Universal Robots URScript: FaiChun_9 Jan_4.script

def Machining1():
  # Default parameters:
  global speed_ms = 0.3
  global speed_rads = 0.75
  global accel_mss = 3
  global accel_radss = 1.2
  global blend_radius_m = 0.0003

  # Add subprograms here
  # Start of main program
  # Program generated by RoboDK v5.6.8 for UR10e on 09/01/2025 17:05:57
  # Using nominal kinematics.
  blend_radius_m = 0.0003
  speed_ms = 0.03
  # set_reference(p[0.335000, -0.060000, 0.000000, 0.000000, 0.000000, 0.000000])
  set_tcp(p[0.000000, 0.000000, 0.252000, 0.000000, 0.000000, 0.000000])
  # Show Tool
  movej([0.372931, -1.100475, -2.621390, -0.990524, 1.570796, 1.943727],accel_radss,speed_rads,0,blend_radius_m)
  movel([0.372931, -1.160560, -2.660288, -0.891541, 1.570796, 1.943727],accel_mss,speed_ms,0,blend_radius_m)
  #SetTool1
  #M_RunCode6
  #SetRPM60000
  speed_ms = 0.03
  #M_RunCode3
  movel([0.372931, -1.188229, -2.675077, -0.849084, 1.570796, 1.943727],accel_mss,speed_ms,0,blend_radius_m)
  speed_ms = 0.003
  movel([0.372931, -1.195517, -2.678710, -0.838162, 1.570796, 1.943727],accel_mss,speed_ms,0,blend_radius_m)
  speed_ms = 0.007
  movel([0.375174, -1.198382, -2.677355, -0.836652, 1.570796, 1.945970],accel_mss,speed_ms,0,blend_radius_m)
  movel([0.377606, -1.200493, -2.676351, -0.835545, 1.570796, 1.948402],accel_mss,speed_ms,0,blend_radius_m)
  movel([0.380241, -1.201847, -2.675704, -0.834837, 1.570796, 1.951037],accel_mss,speed_ms,0,blend_radius_m)
  movel([0.383075, -1.202452, -2.675415, -0.834522, 1.570796, 1.953872],accel_mss,speed_ms,0,blend_radius_m)
  movel([0.386053, -1.202396, -2.675442, -0.834551, 1.570796, 1.956849],accel_mss,speed_ms,0,blend_radius_m)
  movel([0.389105, -1.201761, -2.675746, -0.834882, 1.570796, 1.959901],accel_mss,speed_ms,0,blend_radius_m)
  movel([0.392242, -1.200547, -2.676325, -0.835516, 1.570796, 1.963038],accel_mss,speed_ms,0,blend_radius_m)
  movel([0.395468, -1.198746, -2.677183, -0.836461, 1.570796, 1.966265],accel_mss,speed_ms,0,blend_radius_m)
  movel([0.380728, -1.210997, -2.671282, -0.830110, 1.570796, 1.951524],accel_mss,speed_ms,0,blend_radius_m)
  movel([0.361187, -1.181602, -2.685164, -0.845623, 1.570796, 1.931983],accel_mss,speed_ms,0,blend_radius_m)
  movel([0.362683, -1.180288, -2.685763, -0.846338, 1.570796, 1.933479],accel_mss,speed_ms,0,blend_radius_m)
  movel([0.366731, -1.177285, -2.687125, -0.847980, 1.570796, 1.937528],accel_mss,speed_ms,0,blend_radius_m)
  movel([0.371187, -1.175024, -2.688143, -0.849221, 1.570796, 1.941984],accel_mss,speed_ms,0,blend_radius_m)
  movel([0.375796, -1.173412, -2.688867, -0.850111, 1.570796, 1.946593],accel_mss,speed_ms,0,blend_radius_m)
  movel([0.380308, -1.172343, -2.689344, -0.850701, 1.570796, 1.951104],accel_mss,speed_ms,0,blend_radius_m)
  movel([0.392053, -1.170737, -2.690060, -0.851592, 1.570796, 1.962849],accel_mss,speed_ms,0,blend_radius_m)
  movel([0.402871, -1.169477, -2.690620, -0.852292, 1.570796, 1.973667],accel_mss,speed_ms,0,blend_radius_m)
  movel([0.407062, -1.168614, -2.691003, -0.852772, 1.570796, 1.977858],accel_mss,speed_ms,0,blend_radius_m)
  movel([0.411263, -1.167290, -2.691588, -0.853511, 1.570796, 1.982060],accel_mss,speed_ms,0,blend_radius_m)
  movel([0.415272, -1.165416, -2.692413, -0.854560, 1.570796, 1.986068],accel_mss,speed_ms,0,blend_radius_m)
  movel([0.418891, -1.162891, -2.693519, -0.855978, 1.570796, 1.989688],accel_mss,speed_ms,0,blend_radius_m)
  movel([0.422708, -1.159075, -2.695179, -0.858136, 1.570796, 1.993505],accel_mss,speed_ms,0,blend_radius_m)
  movel([0.424029, -1.157173, -2.696000, -0.859216, 1.570796, 1.994826],accel_mss,speed_ms,0,blend_radius_m)
  movel([0.424957, -1.155274, -2.696817, -0.860298, 1.570796, 1.995753],accel_mss,speed_ms,0,blend_radius_m)
  movel([0.425724, -1.151821, -2.698292, -0.862276, 1.570796, 1.996520],accel_mss,speed_ms,0,blend_radius_m)
  movel([0.425106, -1.149060, -2.699463, -0.863866, 1.570796, 1.995903],accel_mss,speed_ms,0,blend_radius_m)
  movel([0.424036, -1.147738, -2.700021, -0.864630, 1.570796, 1.994833],accel_mss,speed_ms,0,blend_radius_m)
  movel([0.422706, -1.147211, -2.700243, -0.864935, 1.570796, 1.993503],accel_mss,speed_ms,0,blend_radius_m)
  movel([0.421264, -1.147406, -2.700161, -0.864822, 1.570796, 1.992060],accel_mss,speed_ms,0,blend_radius_m)
  movel([0.419851, -1.148255, -2.699803, -0.864331, 1.570796, 1.990647],accel_mss,speed_ms,0,blend_radius_m)
  movel([0.418269, -1.150392, -2.698899, -0.863098, 1.570796, 1.989065],accel_mss,speed_ms,0,blend_radius_m)
  movel([0.416848, -1.152543, -2.697985, -0.861862, 1.570796, 1.987644],accel_mss,speed_ms,0,blend_radius_m)
  movel([0.414611, -1.154776, -2.697030, -0.860583, 1.570796, 1.985407],accel_mss,speed_ms,0,blend_radius_m)
  movel([0.411600, -1.156758, -2.696179, -0.859452, 1.570796, 1.982396],accel_mss,speed_ms,0,blend_radius_m)
  movel([0.408872, -1.157382, -2.695910, -0.859097, 1.570796, 1.979668],accel_mss,speed_ms,0,blend_radius_m)
  movel([0.406625, -1.156830, -2.696148, -0.859411, 1.570796, 1.977422],accel_mss,speed_ms,0,blend_radius_m)
  movel([0.405066, -1.155270, -2.696818, -0.860301, 1.570796, 1.975862],accel_mss,speed_ms,0,blend_radius_m)
  movel([0.404360, -1.152976, -2.697800, -0.861613, 1.570796, 1.975156],accel_mss,speed_ms,0,blend_radius_m)
  movel([0.404684, -1.150222, -2.698971, -0.863196, 1.570796, 1.975481],accel_mss,speed_ms,0,blend_radius_m)
  movel([0.406108, -1.147296, -2.700207, -0.864886, 1.570796, 1.976904],accel_mss,speed_ms,0,blend_radius_m)
  movel([0.408704, -1.144500, -2.701381, -0.866509, 1.570796, 1.979501],accel_mss,speed_ms,0,blend_radius_m)
  movel([0.411321, -1.142589, -2.702178, -0.867622, 1.570796, 1.982118],accel_mss,speed_ms,0,blend_radius_m)
  movel([0.413891, -1.141382, -2.702680, -0.868328, 1.570796, 1.984688],accel_mss,speed_ms,0,blend_radius_m)
  movel([0.416415, -1.140882, -2.702887, -0.868620, 1.570796, 1.987211],accel_mss,speed_ms,0,blend_radius_m)
  movel([0.418874, -1.141102, -2.702796, -0.868491, 1.570796, 1.989670],accel_mss,speed_ms,0,blend_radius_m)
  movel([0.421187, -1.141949, -2.702444, -0.867996, 1.570796, 1.991984],accel_mss,speed_ms,0,blend_radius_m)
  movel([0.423263, -1.143337, -2.701866, -0.867186, 1.570796, 1.994060],accel_mss,speed_ms,0,blend_radius_m)
  movel([0.426702, -1.147727, -2.700026, -0.864636, 1.570796, 1.997499],accel_mss,speed_ms,0,blend_radius_m)
  movel([0.428202, -1.151149, -2.698578, -0.862662, 1.570796, 1.998999],accel_mss,speed_ms,0,blend_radius_m)
  movel([0.429111, -1.154788, -2.697025, -0.860576, 1.570796, 1.999907],accel_mss,speed_ms,0,blend_radius_m)
  movel([0.429435, -1.158639, -2.695367, -0.858383, 1.570796, 2.000231],accel_mss,speed_ms,0,blend_radius_m)
  movel([0.429184, -1.162688, -2.693608, -0.856093, 1.570796, 1.999980],accel_mss,speed_ms,0,blend_radius_m)
  movel([0.428147, -1.166773, -2.691816, -0.853800, 1.570796, 1.998944],accel_mss,speed_ms,0,blend_radius_m)
  movel([0.426123, -1.170732, -2.690063, -0.851595, 1.570796, 1.996919],accel_mss,speed_ms,0,blend_radius_m)
  movel([0.423112, -1.174570, -2.688347, -0.849472, 1.570796, 1.993908],accel_mss,speed_ms,0,blend_radius_m)
  movel([0.419124, -1.178294, -2.686668, -0.847427, 1.570796, 1.989921],accel_mss,speed_ms,0,blend_radius_m)
  movel([0.415165, -1.181134, -2.685378, -0.845877, 1.570796, 1.985962],accel_mss,speed_ms,0,blend_radius_m)
  movel([0.411168, -1.183199, -2.684434, -0.844756, 1.570796, 1.981965],accel_mss,speed_ms,0,blend_radius_m)
  movel([0.407228, -1.184627, -2.683779, -0.843983, 1.570796, 1.978024],accel_mss,speed_ms,0,blend_radius_m)
  movel([0.403450, -1.185553, -2.683353, -0.843483, 1.570796, 1.974246],accel_mss,speed_ms,0,blend_radius_m)
  movel([0.394479, -1.186696, -2.682826, -0.842867, 1.570796, 1.965275],accel_mss,speed_ms,0,blend_radius_m)
  movel([0.385975, -1.187888, -2.682274, -0.842226, 1.570796, 1.956771],accel_mss,speed_ms,0,blend_radius_m)
  movel([0.382534, -1.188768, -2.681867, -0.841754, 1.570796, 1.953330],accel_mss,speed_ms,0,blend_radius_m)
  movel([0.379011, -1.190092, -2.681251, -0.841046, 1.570796, 1.949807],accel_mss,speed_ms,0,blend_radius_m)
  movel([0.375525, -1.191944, -2.680387, -0.840058, 1.570796, 1.946321],accel_mss,speed_ms,0,blend_radius_m)
  movel([0.372203, -1.194411, -2.679231, -0.838747, 1.570796, 1.942999],accel_mss,speed_ms,0,blend_radius_m)
  movel([0.372931, -1.195517, -2.678710, -0.838162, 1.570796, 1.943727],accel_mss,speed_ms,0,blend_radius_m)
  speed_ms = 0.003
  movel([0.372931, -1.188229, -2.675077, -0.849084, 1.570796, 1.943727],accel_mss,speed_ms,0,blend_radius_m)
  speed_ms = 0.03
  movel([0.372931, -1.160560, -2.660288, -0.891541, 1.570796, 1.943727],accel_mss,speed_ms,0,blend_radius_m)
  #M_RunCode9
  movel([0.396562, -1.185032, -2.648957, -0.878400, 1.570796, 1.967359],accel_mss,speed_ms,0,blend_radius_m)
  #M_RunCode3
  movel([0.396562, -1.212507, -2.663422, -0.836459, 1.570796, 1.967359],accel_mss,speed_ms,0,blend_radius_m)
  speed_ms = 0.003
  movel([0.396562, -1.219730, -2.666973, -0.825686, 1.570796, 1.967359],accel_mss,speed_ms,0,blend_radius_m)
  speed_ms = 0.007
  movel([0.404177, -1.212524, -2.670535, -0.829330, 1.570796, 1.974973],accel_mss,speed_ms,0,blend_radius_m)
  movel([0.415586, -1.202971, -2.675166, -0.834252, 1.570796, 1.986383],accel_mss,speed_ms,0,blend_radius_m)
  movel([0.427444, -1.193807, -2.679515, -0.839067, 1.570796, 1.998240],accel_mss,speed_ms,0,blend_radius_m)
  movel([0.436211, -1.187874, -2.682281, -0.842234, 1.570796, 2.007007],accel_mss,speed_ms,0,blend_radius_m)
  movel([0.439450, -1.186181, -2.683064, -0.843145, 1.570796, 2.010246],accel_mss,speed_ms,0,blend_radius_m)
  movel([0.441984, -1.185395, -2.683426, -0.843569, 1.570796, 2.012781],accel_mss,speed_ms,0,blend_radius_m)
  movel([0.443806, -1.185518, -2.683369, -0.843502, 1.570796, 2.014603],accel_mss,speed_ms,0,blend_radius_m)
  movel([0.444914, -1.186554, -2.682891, -0.842944, 1.570796, 2.015710],accel_mss,speed_ms,0,blend_radius_m)
  movel([0.445184, -1.188242, -2.682110, -0.842036, 1.570796, 2.015980],accel_mss,speed_ms,0,blend_radius_m)
  movel([0.444497, -1.190341, -2.681135, -0.840912, 1.570796, 2.015293],accel_mss,speed_ms,0,blend_radius_m)
  movel([0.442860, -1.192839, -2.679968, -0.839581, 1.570796, 2.013656],accel_mss,speed_ms,0,blend_radius_m)
  movel([0.440283, -1.195736, -2.678607, -0.838046, 1.570796, 2.011079],accel_mss,speed_ms,0,blend_radius_m)
  movel([0.432369, -1.203009, -2.675148, -0.834232, 1.570796, 2.003165],accel_mss,speed_ms,0,blend_radius_m)
  movel([0.420879, -1.212434, -2.670579, -0.829376, 1.570796, 1.991675],accel_mss,speed_ms,0,blend_radius_m)
  movel([0.409297, -1.221297, -2.666191, -0.824901, 1.570796, 1.980094],accel_mss,speed_ms,0,blend_radius_m)
  movel([0.400914, -1.226977, -2.663332, -0.822080, 1.570796, 1.971711],accel_mss,speed_ms,0,blend_radius_m)
  movel([0.397832, -1.228606, -2.662505, -0.821278, 1.570796, 1.968628],accel_mss,speed_ms,0,blend_radius_m)
  movel([0.395403, -1.229390, -2.662106, -0.820893, 1.570796, 1.966199],accel_mss,speed_ms,0,blend_radius_m)
  movel([0.393621, -1.229327, -2.662138, -0.820924, 1.570796, 1.964417],accel_mss,speed_ms,0,blend_radius_m)
  movel([0.392480, -1.228419, -2.662600, -0.821370, 1.570796, 1.963276],accel_mss,speed_ms,0,blend_radius_m)
  movel([0.392118, -1.226877, -2.663382, -0.822130, 1.570796, 1.962915],accel_mss,speed_ms,0,blend_radius_m)
  movel([0.392674, -1.224917, -2.664373, -0.823099, 1.570796, 1.963470],accel_mss,speed_ms,0,blend_radius_m)
  movel([0.394153, -1.222536, -2.665570, -0.824283, 1.570796, 1.964950],accel_mss,speed_ms,0,blend_radius_m)
  movel([0.396562, -1.219730, -2.666973, -0.825686, 1.570796, 1.967359],accel_mss,speed_ms,0,blend_radius_m)
  speed_ms = 0.003
  movel([0.396562, -1.212507, -2.663422, -0.836459, 1.570796, 1.967359],accel_mss,speed_ms,0,blend_radius_m)
  speed_ms = 0.03
  movel([0.396562, -1.185032, -2.648957, -0.878400, 1.570796, 1.967359],accel_mss,speed_ms,0,blend_radius_m)
  #M_RunCode9
  movel([0.389349, -1.187940, -2.647569, -0.876881, 1.570796, 1.960145],accel_mss,speed_ms,0,blend_radius_m)
  #M_RunCode3
  movel([0.389349, -1.215389, -2.661996, -0.835005, 1.570796, 1.960145],accel_mss,speed_ms,0,blend_radius_m)
  speed_ms = 0.003
  movel([0.389349, -1.222603, -2.665537, -0.824249, 1.570796, 1.960145],accel_mss,speed_ms,0,blend_radius_m)
  speed_ms = 0.007
  movel([0.389682, -1.219825, -2.666926, -0.825638, 1.570796, 1.960478],accel_mss,speed_ms,0,blend_radius_m)
  movel([0.390483, -1.216852, -2.668402, -0.827134, 1.570796, 1.961280],accel_mss,speed_ms,0,blend_radius_m)
  movel([0.391770, -1.213727, -2.669944, -0.828718, 1.570796, 1.962567],accel_mss,speed_ms,0,blend_radius_m)
  movel([0.393551, -1.210442, -2.671553, -0.830394, 1.570796, 1.964348],accel_mss,speed_ms,0,blend_radius_m)
  movel([0.395827, -1.207003, -2.673224, -0.832162, 1.570796, 1.966623],accel_mss,speed_ms,0,blend_radius_m)
  movel([0.398587, -1.203463, -2.674930, -0.833996, 1.570796, 1.969383],accel_mss,speed_ms,0,blend_radius_m)
  movel([0.401818, -1.199899, -2.676634, -0.835856, 1.570796, 1.972615],accel_mss,speed_ms,0,blend_radius_m)
  movel([0.405529, -1.196306, -2.678338, -0.837745, 1.570796, 1.976325],accel_mss,speed_ms,0,blend_radius_m)
  movel([0.409718, -1.192689, -2.680039, -0.839661, 1.570796, 1.980515],accel_mss,speed_ms,0,blend_radius_m)
  movel([0.414077, -1.189311, -2.681615, -0.841464, 1.570796, 1.984873],accel_mss,speed_ms,0,blend_radius_m)
  movel([0.418282, -1.186435, -2.682946, -0.843008, 1.570796, 1.989078],accel_mss,speed_ms,0,blend_radius_m)
  movel([0.422334, -1.184063, -2.684038, -0.844288, 1.570796, 1.993130],accel_mss,speed_ms,0,blend_radius_m)
  movel([0.426217, -1.182209, -2.684887, -0.845293, 1.570796, 1.997013],accel_mss,speed_ms,0,blend_radius_m)
  movel([0.429866, -1.180871, -2.685498, -0.846020, 1.570796, 2.000662],accel_mss,speed_ms,0,blend_radius_m)
  movel([0.433215, -1.180048, -2.685872, -0.846468, 1.570796, 2.004011],accel_mss,speed_ms,0,blend_radius_m)
  movel([0.436251, -1.179750, -2.686008, -0.846632, 1.570796, 2.007047],accel_mss,speed_ms,0,blend_radius_m)
  movel([0.438978, -1.179968, -2.685909, -0.846512, 1.570796, 2.009774],accel_mss,speed_ms,0,blend_radius_m)
  movel([0.441366, -1.180667, -2.685591, -0.846131, 1.570796, 2.012162],accel_mss,speed_ms,0,blend_radius_m)
  movel([0.443394, -1.181812, -2.685068, -0.845508, 1.570796, 2.014190],accel_mss,speed_ms,0,blend_radius_m)
  movel([0.445058, -1.183393, -2.684345, -0.844651, 1.570796, 2.015855],accel_mss,speed_ms,0,blend_radius_m)
  movel([0.446358, -1.185415, -2.683416, -0.843557, 1.570796, 2.017155],accel_mss,speed_ms,0,blend_radius_m)
  movel([0.447245, -1.187753, -2.682337, -0.842299, 1.570796, 2.018041],accel_mss,speed_ms,0,blend_radius_m)
  movel([0.447665, -1.190296, -2.681156, -0.840937, 1.570796, 2.018461],accel_mss,speed_ms,0,blend_radius_m)
  movel([0.447622, -1.193039, -2.679875, -0.839475, 1.570796, 2.018418],accel_mss,speed_ms,0,blend_radius_m)
  movel([0.447118, -1.195977, -2.678493, -0.837919, 1.570796, 2.017915],accel_mss,speed_ms,0,blend_radius_m)
  movel([0.446145, -1.199069, -2.677029, -0.836291, 1.570796, 2.016941],accel_mss,speed_ms,0,blend_radius_m)
  movel([0.444689, -1.202271, -2.675502, -0.834616, 1.570796, 2.015486],accel_mss,speed_ms,0,blend_radius_m)
  movel([0.442760, -1.205576, -2.673913, -0.832899, 1.570796, 2.013556],accel_mss,speed_ms,0,blend_radius_m)
  movel([0.440355, -1.208991, -2.672259, -0.831138, 1.570796, 2.011152],accel_mss,speed_ms,0,blend_radius_m)
  movel([0.437506, -1.212440, -2.670576, -0.829373, 1.570796, 2.008302],accel_mss,speed_ms,0,blend_radius_m)
  movel([0.434240, -1.215858, -2.668894, -0.827637, 1.570796, 2.005036],accel_mss,speed_ms,0,blend_radius_m)
  movel([0.430553, -1.219251, -2.667212, -0.825926, 1.570796, 2.001350],accel_mss,speed_ms,0,blend_radius_m)
  movel([0.426454, -1.222616, -2.665530, -0.824243, 1.570796, 1.997250],accel_mss,speed_ms,0,blend_radius_m)
  movel([0.422240, -1.225730, -2.663962, -0.822696, 1.570796, 1.993036],accel_mss,speed_ms,0,blend_radius_m)
  movel([0.418217, -1.228354, -2.662633, -0.821402, 1.570796, 1.989014],accel_mss,speed_ms,0,blend_radius_m)
  movel([0.414369, -1.230502, -2.661539, -0.820348, 1.570796, 1.985165],accel_mss,speed_ms,0,blend_radius_m)
  movel([0.410696, -1.232176, -2.660682, -0.819531, 1.570796, 1.981492],accel_mss,speed_ms,0,blend_radius_m)
  movel([0.407244, -1.233389, -2.660060, -0.818941, 1.570796, 1.978040],accel_mss,speed_ms,0,blend_radius_m)
  movel([0.404067, -1.234145, -2.659671, -0.818573, 1.570796, 1.974863],accel_mss,speed_ms,0,blend_radius_m)
  movel([0.401160, -1.234451, -2.659513, -0.818425, 1.570796, 1.971956],accel_mss,speed_ms,0,blend_radius_m)
  movel([0.398519, -1.234302, -2.659590, -0.818497, 1.570796, 1.969315],accel_mss,speed_ms,0,blend_radius_m)
  movel([0.396172, -1.233724, -2.659887, -0.818778, 1.570796, 1.966969],accel_mss,speed_ms,0,blend_radius_m)
  movel([0.394146, -1.232747, -2.660389, -0.819253, 1.570796, 1.964942],accel_mss,speed_ms,0,blend_radius_m)
  movel([0.392438, -1.231366, -2.661097, -0.819926, 1.570796, 1.963234],accel_mss,speed_ms,0,blend_radius_m)
  movel([0.391047, -1.229578, -2.662010, -0.820801, 1.570796, 1.961843],accel_mss,speed_ms,0,blend_radius_m)
  movel([0.390035, -1.227475, -2.663079, -0.821835, 1.570796, 1.960831],accel_mss,speed_ms,0,blend_radius_m)
  movel([0.389467, -1.225152, -2.664254, -0.822982, 1.570796, 1.960264],accel_mss,speed_ms,0,blend_radius_m)
  movel([0.389349, -1.222603, -2.665537, -0.824249, 1.570796, 1.960145],accel_mss,speed_ms,0,blend_radius_m)
  speed_ms = 0.003
  movel([0.389349, -1.215389, -2.661996, -0.835005, 1.570796, 1.960145],accel_mss,speed_ms,0,blend_radius_m)
  speed_ms = 0.03
  movel([0.389349, -1.187940, -2.647569, -0.876881, 1.570796, 1.960145],accel_mss,speed_ms,0,blend_radius_m)
  #M_RunCode9
  movel([0.511389, -1.442779, -2.486051, -0.783559, 1.570796, 2.082185],accel_mss,speed_ms,0,blend_radius_m)
  #M_RunCode3
  movel([0.511389, -1.466101, -2.497203, -0.749085, 1.570796, 2.082185],accel_mss,speed_ms,0,blend_radius_m)
  speed_ms = 0.003
  movel([0.511389, -1.472126, -2.499919, -0.740344, 1.570796, 2.082185],accel_mss,speed_ms,0,blend_radius_m)
  speed_ms = 0.007
  movel([0.512510, -1.471509, -2.500439, -0.740441, 1.570796, 2.083306],accel_mss,speed_ms,0,blend_radius_m)
  movel([0.515465, -1.470227, -2.501517, -0.740644, 1.570796, 2.086261],accel_mss,speed_ms,0,blend_radius_m)
  movel([0.518585, -1.469544, -2.502091, -0.740754, 1.570796, 2.089381],accel_mss,speed_ms,0,blend_radius_m)
  movel([0.521721, -1.469336, -2.502266, -0.740787, 1.570796, 2.092517],accel_mss,speed_ms,0,blend_radius_m)
  movel([0.524727, -1.469486, -2.502140, -0.740763, 1.570796, 2.095523],accel_mss,speed_ms,0,blend_radius_m)
  movel([0.532413, -1.470666, -2.501149, -0.740574, 1.570796, 2.103210],accel_mss,speed_ms,0,blend_radius_m)
  movel([0.539462, -1.471881, -2.500125, -0.740383, 1.570796, 2.110258],accel_mss,speed_ms,0,blend_radius_m)
  movel([0.542231, -1.472091, -2.499948, -0.740350, 1.570796, 2.113027],accel_mss,speed_ms,0,blend_radius_m)
  movel([0.545054, -1.471987, -2.500036, -0.740366, 1.570796, 2.115850],accel_mss,speed_ms,0,blend_radius_m)
  movel([0.547810, -1.471472, -2.500470, -0.740447, 1.570796, 2.118606],accel_mss,speed_ms,0,blend_radius_m)
  movel([0.550379, -1.470448, -2.501332, -0.740609, 1.570796, 2.121175],accel_mss,speed_ms,0,blend_radius_m)
  movel([0.553203, -1.468592, -2.502890, -0.740907, 1.570796, 2.123999],accel_mss,speed_ms,0,blend_radius_m)
  movel([0.554237, -1.467561, -2.503753, -0.741075, 1.570796, 2.125033],accel_mss,speed_ms,0,blend_radius_m)
  movel([0.555022, -1.466457, -2.504675, -0.741257, 1.570796, 2.125818],accel_mss,speed_ms,0,blend_radius_m)
  movel([0.555859, -1.464286, -2.506484, -0.741620, 1.570796, 2.126655],accel_mss,speed_ms,0,blend_radius_m)
  movel([0.555749, -1.462318, -2.508116, -0.741955, 1.570796, 2.126546],accel_mss,speed_ms,0,blend_radius_m)
  movel([0.555208, -1.461229, -2.509018, -0.742143, 1.570796, 2.126004],accel_mss,speed_ms,0,blend_radius_m)
  movel([0.554422, -1.460619, -2.509521, -0.742249, 1.570796, 2.125218],accel_mss,speed_ms,0,blend_radius_m)
  movel([0.553489, -1.460476, -2.509639, -0.742274, 1.570796, 2.124285],accel_mss,speed_ms,0,blend_radius_m)
  movel([0.552509, -1.460776, -2.509392, -0.742221, 1.570796, 2.123306],accel_mss,speed_ms,0,blend_radius_m)
  movel([0.551284, -1.461908, -2.508456, -0.742025, 1.570796, 2.122080],accel_mss,speed_ms,0,blend_radius_m)
  movel([0.550160, -1.463080, -2.507485, -0.741824, 1.570796, 2.120957],accel_mss,speed_ms,0,blend_radius_m)
  movel([0.548506, -1.464159, -2.506589, -0.741641, 1.570796, 2.119302],accel_mss,speed_ms,0,blend_radius_m)
  movel([0.546387, -1.464918, -2.505958, -0.741513, 1.570796, 2.117183],accel_mss,speed_ms,0,blend_radius_m)
  movel([0.544590, -1.464817, -2.506042, -0.741530, 1.570796, 2.115386],accel_mss,speed_ms,0,blend_radius_m)
  movel([0.543223, -1.464011, -2.506712, -0.741666, 1.570796, 2.114019],accel_mss,speed_ms,0,blend_radius_m)
  movel([0.542400, -1.462654, -2.507838, -0.741897, 1.570796, 2.113196],accel_mss,speed_ms,0,blend_radius_m)
  movel([0.542203, -1.460966, -2.509235, -0.742188, 1.570796, 2.112999],accel_mss,speed_ms,0,blend_radius_m)
  movel([0.542704, -1.459169, -2.510717, -0.742503, 1.570796, 2.113500],accel_mss,speed_ms,0,blend_radius_m)
  movel([0.543921, -1.457473, -2.512111, -0.742805, 1.570796, 2.114717],accel_mss,speed_ms,0,blend_radius_m)
  movel([0.545862, -1.456097, -2.513239, -0.743053, 1.570796, 2.116658],accel_mss,speed_ms,0,blend_radius_m)
  movel([0.547718, -1.455322, -2.513873, -0.743194, 1.570796, 2.118514],accel_mss,speed_ms,0,blend_radius_m)
  movel([0.549468, -1.455012, -2.514126, -0.743251, 1.570796, 2.120264],accel_mss,speed_ms,0,blend_radius_m)
  movel([0.551108, -1.455170, -2.513997, -0.743222, 1.570796, 2.121904],accel_mss,speed_ms,0,blend_radius_m)
  movel([0.552636, -1.455794, -2.513487, -0.743108, 1.570796, 2.123433],accel_mss,speed_ms,0,blend_radius_m)
  movel([0.554006, -1.456805, -2.512659, -0.742925, 1.570796, 2.124803],accel_mss,speed_ms,0,blend_radius_m)
  movel([0.555173, -1.458135, -2.511567, -0.742687, 1.570796, 2.125970],accel_mss,speed_ms,0,blend_radius_m)
  movel([0.556897, -1.461726, -2.508606, -0.742056, 1.570796, 2.127693],accel_mss,speed_ms,0,blend_radius_m)
  movel([0.557498, -1.464304, -2.506469, -0.741616, 1.570796, 2.128294],accel_mss,speed_ms,0,blend_radius_m)
  movel([0.557707, -1.466914, -2.504293, -0.741181, 1.570796, 2.128503],accel_mss,speed_ms,0,blend_radius_m)
  movel([0.557526, -1.469558, -2.502079, -0.740751, 1.570796, 2.128322],accel_mss,speed_ms,0,blend_radius_m)
  movel([0.556957, -1.472236, -2.499826, -0.740327, 1.570796, 2.127754],accel_mss,speed_ms,0,blend_radius_m)
  movel([0.555888, -1.474796, -2.497662, -0.739932, 1.570796, 2.126684],accel_mss,speed_ms,0,blend_radius_m)
  movel([0.554191, -1.477097, -2.495707, -0.739585, 1.570796, 2.124987],accel_mss,speed_ms,0,blend_radius_m)
  movel([0.551872, -1.479141, -2.493964, -0.739284, 1.570796, 2.122669],accel_mss,speed_ms,0,blend_radius_m)
  movel([0.548934, -1.480933, -2.492431, -0.739025, 1.570796, 2.119730],accel_mss,speed_ms,0,blend_radius_m)
  movel([0.546095, -1.482138, -2.491397, -0.738854, 1.570796, 2.116892],accel_mss,speed_ms,0,blend_radius_m)
  movel([0.543309, -1.482807, -2.490821, -0.738760, 1.570796, 2.114105],accel_mss,speed_ms,0,blend_radius_m)
  movel([0.540622, -1.483053, -2.490610, -0.738726, 1.570796, 2.111419],accel_mss,speed_ms,0,blend_radius_m)
  movel([0.538093, -1.482982, -2.490671, -0.738736, 1.570796, 2.108889],accel_mss,speed_ms,0,blend_radius_m)
  movel([0.532193, -1.482083, -2.491443, -0.738862, 1.570796, 2.102990],accel_mss,speed_ms,0,blend_radius_m)
  movel([0.526586, -1.481294, -2.492121, -0.738974, 1.570796, 2.097382],accel_mss,speed_ms,0,blend_radius_m)
  movel([0.524266, -1.481248, -2.492160, -0.738981, 1.570796, 2.095063],accel_mss,speed_ms,0,blend_radius_m)
  movel([0.521845, -1.481490, -2.491953, -0.738946, 1.570796, 2.092642],accel_mss,speed_ms,0,blend_radius_m)
  movel([0.519382, -1.482109, -2.491422, -0.738859, 1.570796, 2.090178],accel_mss,speed_ms,0,blend_radius_m)
  movel([0.516949, -1.483187, -2.490495, -0.738707, 1.570796, 2.087746],accel_mss,speed_ms,0,blend_radius_m)
  movel([0.517290, -1.484097, -2.489711, -0.738581, 1.570796, 2.088086],accel_mss,speed_ms,0,blend_radius_m)
  movel([0.518405, -1.486522, -2.487616, -0.738252, 1.570796, 2.089201],accel_mss,speed_ms,0,blend_radius_m)
  movel([0.519736, -1.488456, -2.485938, -0.737995, 1.570796, 2.090533],accel_mss,speed_ms,0,blend_radius_m)
  movel([0.521285, -1.489897, -2.484684, -0.737808, 1.570796, 2.092082],accel_mss,speed_ms,0,blend_radius_m)
  movel([0.523056, -1.490852, -2.483852, -0.737686, 1.570796, 2.093852],accel_mss,speed_ms,0,blend_radius_m)
  movel([0.524991, -1.491371, -2.483399, -0.737620, 1.570796, 2.095787],accel_mss,speed_ms,0,blend_radius_m)
  movel([0.527041, -1.491500, -2.483286, -0.737603, 1.570796, 2.097838],accel_mss,speed_ms,0,blend_radius_m)
  movel([0.529210, -1.491241, -2.483512, -0.737636, 1.570796, 2.100007],accel_mss,speed_ms,0,blend_radius_m)
  movel([0.531500, -1.490592, -2.484078, -0.737719, 1.570796, 2.102296],accel_mss,speed_ms,0,blend_radius_m)
  movel([0.520553, -1.496378, -2.479005, -0.737006, 1.570796, 2.091350],accel_mss,speed_ms,0,blend_radius_m)
  movel([0.511389, -1.472126, -2.499919, -0.740344, 1.570796, 2.082185],accel_mss,speed_ms,0,blend_radius_m)
  speed_ms = 0.003
  movel([0.511389, -1.466101, -2.497203, -0.749085, 1.570796, 2.082185],accel_mss,speed_ms,0,blend_radius_m)
  speed_ms = 0.03
  movel([0.511389, -1.442779, -2.486051, -0.783559, 1.570796, 2.082185],accel_mss,speed_ms,0,blend_radius_m)
  #M_RunCode9
  movel([0.528462, -1.467084, -2.466023, -0.779282, 1.570796, 2.099259],accel_mss,speed_ms,0,blend_radius_m)
  #M_RunCode3
  movel([0.528462, -1.489892, -2.476890, -0.745607, 1.570796, 2.099259],accel_mss,speed_ms,0,blend_radius_m)
  speed_ms = 0.003
  movel([0.528462, -1.495777, -2.479534, -0.737078, 1.570796, 2.099259],accel_mss,speed_ms,0,blend_radius_m)
  speed_ms = 0.007
  movel([0.530510, -1.495038, -2.480185, -0.737166, 1.570796, 2.101306],accel_mss,speed_ms,0,blend_radius_m)
  movel([0.532280, -1.495118, -2.480114, -0.737157, 1.570796, 2.103076],accel_mss,speed_ms,0,blend_radius_m)
  movel([0.533639, -1.495877, -2.479446, -0.737066, 1.570796, 2.104435],accel_mss,speed_ms,0,blend_radius_m)
  movel([0.534453, -1.497172, -2.478305, -0.736912, 1.570796, 2.105249],accel_mss,speed_ms,0,blend_radius_m)
  movel([0.534648, -1.498784, -2.476880, -0.736725, 1.570796, 2.105445],accel_mss,speed_ms,0,blend_radius_m)
  movel([0.534160, -1.500498, -2.475360, -0.736531, 1.570796, 2.104956],accel_mss,speed_ms,0,blend_radius_m)
  movel([0.532994, -1.502101, -2.473935, -0.736353, 1.570796, 2.103791],accel_mss,speed_ms,0,blend_radius_m)
  movel([0.531163, -1.503383, -2.472792, -0.736214, 1.570796, 2.101959],accel_mss,speed_ms,0,blend_radius_m)
  movel([0.529477, -1.504055, -2.472192, -0.736142, 1.570796, 2.100273],accel_mss,speed_ms,0,blend_radius_m)
  movel([0.528093, -1.504217, -2.472047, -0.736125, 1.570796, 2.098889],accel_mss,speed_ms,0,blend_radius_m)
  movel([0.526667, -1.504492, -2.471802, -0.736095, 1.570796, 2.097463],accel_mss,speed_ms,0,blend_radius_m)
  movel([0.525860, -1.505120, -2.471240, -0.736029, 1.570796, 2.096656],accel_mss,speed_ms,0,blend_radius_m)
  movel([0.525333, -1.506016, -2.470437, -0.735936, 1.570796, 2.096129],accel_mss,speed_ms,0,blend_radius_m)
  movel([0.525125, -1.507024, -2.469533, -0.735833, 1.570796, 2.095921],accel_mss,speed_ms,0,blend_radius_m)
  movel([0.525285, -1.507983, -2.468670, -0.735736, 1.570796, 2.096081],accel_mss,speed_ms,0,blend_radius_m)
  movel([0.525864, -1.509059, -2.467701, -0.735629, 1.570796, 2.096660],accel_mss,speed_ms,0,blend_radius_m)
  movel([0.526729, -1.509863, -2.466976, -0.735550, 1.570796, 2.097525],accel_mss,speed_ms,0,blend_radius_m)
  movel([0.527878, -1.510398, -2.466493, -0.735498, 1.570796, 2.098674],accel_mss,speed_ms,0,blend_radius_m)
  movel([0.529312, -1.510665, -2.466252, -0.735472, 1.570796, 2.100108],accel_mss,speed_ms,0,blend_radius_m)
  movel([0.530946, -1.510650, -2.466265, -0.735474, 1.570796, 2.101742],accel_mss,speed_ms,0,blend_radius_m)
  movel([0.532698, -1.510340, -2.466546, -0.735504, 1.570796, 2.103494],accel_mss,speed_ms,0,blend_radius_m)
  movel([0.534569, -1.509731, -2.467095, -0.735563, 1.570796, 2.105365],accel_mss,speed_ms,0,blend_radius_m)
  movel([0.536560, -1.508826, -2.467911, -0.735652, 1.570796, 2.107356],accel_mss,speed_ms,0,blend_radius_m)
  movel([0.539707, -1.506789, -2.469743, -0.735857, 1.570796, 2.110503],accel_mss,speed_ms,0,blend_radius_m)
  movel([0.542284, -1.504194, -2.472068, -0.736127, 1.570796, 2.113081],accel_mss,speed_ms,0,blend_radius_m)
  movel([0.543329, -1.502697, -2.473404, -0.736288, 1.570796, 2.114126],accel_mss,speed_ms,0,blend_radius_m)
  movel([0.544167, -1.501077, -2.474846, -0.736466, 1.570796, 2.114963],accel_mss,speed_ms,0,blend_radius_m)
  movel([0.545226, -1.497469, -2.478042, -0.736878, 1.570796, 2.116022],accel_mss,speed_ms,0,blend_radius_m)
  movel([0.545348, -1.493463, -2.481567, -0.737358, 1.570796, 2.116144],accel_mss,speed_ms,0,blend_radius_m)
  movel([0.544406, -1.489161, -2.485325, -0.737903, 1.570796, 2.115203],accel_mss,speed_ms,0,blend_radius_m)
  movel([0.561462, -1.480483, -2.492816, -0.739090, 1.570796, 2.132258],accel_mss,speed_ms,0,blend_radius_m)
  movel([0.567091, -1.499193, -2.476518, -0.736678, 1.570796, 2.137887],accel_mss,speed_ms,0,blend_radius_m)
  movel([0.556161, -1.504596, -2.471708, -0.736084, 1.570796, 2.126957],accel_mss,speed_ms,0,blend_radius_m)
  movel([0.558546, -1.502603, -2.473488, -0.736298, 1.570796, 2.129343],accel_mss,speed_ms,0,blend_radius_m)
  movel([0.560525, -1.500138, -2.475680, -0.736571, 1.570796, 2.131322],accel_mss,speed_ms,0,blend_radius_m)
  movel([0.561994, -1.497317, -2.478177, -0.736895, 1.570796, 2.132790],accel_mss,speed_ms,0,blend_radius_m)
  movel([0.562847, -1.494261, -2.480867, -0.737261, 1.570796, 2.133644],accel_mss,speed_ms,0,blend_radius_m)
  movel([0.563020, -1.491086, -2.483647, -0.737656, 1.570796, 2.133816],accel_mss,speed_ms,0,blend_radius_m)
  movel([0.562438, -1.487919, -2.486405, -0.738066, 1.570796, 2.133234],accel_mss,speed_ms,0,blend_radius_m)
  movel([0.549925, -1.494218, -2.480905, -0.737266, 1.570796, 2.120721],accel_mss,speed_ms,0,blend_radius_m)
  movel([0.550757, -1.498036, -2.477542, -0.736812, 1.570796, 2.121553],accel_mss,speed_ms,0,blend_radius_m)
  movel([0.550849, -1.502030, -2.473998, -0.736361, 1.570796, 2.121645],accel_mss,speed_ms,0,blend_radius_m)
  movel([0.550098, -1.505982, -2.470467, -0.735940, 1.570796, 2.120894],accel_mss,speed_ms,0,blend_radius_m)
  movel([0.549366, -1.507863, -2.468778, -0.735748, 1.570796, 2.120163],accel_mss,speed_ms,0,blend_radius_m)
  movel([0.548397, -1.509680, -2.467141, -0.735568, 1.570796, 2.119193],accel_mss,speed_ms,0,blend_radius_m)
  movel([0.547173, -1.511379, -2.465606, -0.735404, 1.570796, 2.117970],accel_mss,speed_ms,0,blend_radius_m)
  movel([0.545678, -1.512905, -2.464223, -0.735261, 1.570796, 2.116474],accel_mss,speed_ms,0,blend_radius_m)
  movel([0.543913, -1.514258, -2.462994, -0.735138, 1.570796, 2.114709],accel_mss,speed_ms,0,blend_radius_m)
  movel([0.541875, -1.515443, -2.461914, -0.735032, 1.570796, 2.112671],accel_mss,speed_ms,0,blend_radius_m)
  movel([0.539753, -1.516377, -2.461062, -0.734950, 1.570796, 2.110549],accel_mss,speed_ms,0,blend_radius_m)
  movel([0.537729, -1.516976, -2.460515, -0.734898, 1.570796, 2.108526],accel_mss,speed_ms,0,blend_radius_m)
  movel([0.535801, -1.517243, -2.460271, -0.734875, 1.570796, 2.106597],accel_mss,speed_ms,0,blend_radius_m)
  movel([0.533968, -1.517180, -2.460329, -0.734880, 1.570796, 2.104764],accel_mss,speed_ms,0,blend_radius_m)
  movel([0.530685, -1.516269, -2.461161, -0.734959, 1.570796, 2.101481],accel_mss,speed_ms,0,blend_radius_m)
  movel([0.527969, -1.514459, -2.462811, -0.735120, 1.570796, 2.098766],accel_mss,speed_ms,0,blend_radius_m)
  movel([0.525859, -1.511972, -2.465069, -0.735348, 1.570796, 2.096656],accel_mss,speed_ms,0,blend_radius_m)
  movel([0.524389, -1.509041, -2.467717, -0.735630, 1.570796, 2.095185],accel_mss,speed_ms,0,blend_radius_m)
  movel([0.523831, -1.506790, -2.469742, -0.735856, 1.570796, 2.094627],accel_mss,speed_ms,0,blend_radius_m)
  movel([0.523699, -1.504279, -2.471992, -0.736118, 1.570796, 2.094495],accel_mss,speed_ms,0,blend_radius_m)
  movel([0.524054, -1.501716, -2.474278, -0.736395, 1.570796, 2.094850],accel_mss,speed_ms,0,blend_radius_m)
  movel([0.524960, -1.499317, -2.476408, -0.736664, 1.570796, 2.095756],accel_mss,speed_ms,0,blend_radius_m)
  movel([0.526426, -1.497272, -2.478216, -0.736901, 1.570796, 2.097222],accel_mss,speed_ms,0,blend_radius_m)
  movel([0.528462, -1.495777, -2.479534, -0.737078, 1.570796, 2.099259],accel_mss,speed_ms,0,blend_radius_m)
  speed_ms = 0.003
  movel([0.528462, -1.489892, -2.476890, -0.745607, 1.570796, 2.099259],accel_mss,speed_ms,0,blend_radius_m)
  speed_ms = 0.03
  movel([0.528462, -1.467084, -2.466023, -0.779282, 1.570796, 2.099259],accel_mss,speed_ms,0,blend_radius_m)
  #M_RunCode9
  movel([0.538901, -1.367315, -2.542780, -0.802295, 1.570796, 2.109697],accel_mss,speed_ms,0,blend_radius_m)
  #M_RunCode3
  movel([0.538901, -1.392148, -2.554861, -0.765381, 1.570796, 2.109697],accel_mss,speed_ms,0,blend_radius_m)
  speed_ms = 0.003
  movel([0.538901, -1.398590, -2.557808, -0.755990, 1.570796, 2.109697],accel_mss,speed_ms,0,blend_radius_m)
  speed_ms = 0.007
  movel([0.535431, -1.399095, -2.557438, -0.755855, 1.570796, 2.106227],accel_mss,speed_ms,0,blend_radius_m)
  movel([0.532084, -1.398897, -2.557584, -0.755908, 1.570796, 2.102881],accel_mss,speed_ms,0,blend_radius_m)
  movel([0.528922, -1.398122, -2.558151, -0.756116, 1.570796, 2.099719],accel_mss,speed_ms,0,blend_radius_m)
  movel([0.526015, -1.396890, -2.559051, -0.756448, 1.570796, 2.096812],accel_mss,speed_ms,0,blend_radius_m)
  movel([0.523439, -1.395316, -2.560198, -0.756875, 1.570796, 2.094235],accel_mss,speed_ms,0,blend_radius_m)
  movel([0.525518, -1.391374, -2.563054, -0.757961, 1.570796, 2.096314],accel_mss,speed_ms,0,blend_radius_m)
  movel([0.528755, -1.387196, -2.566056, -0.759137, 1.570796, 2.099551],accel_mss,speed_ms,0,blend_radius_m)
  movel([0.532819, -1.383159, -2.568934, -0.760297, 1.570796, 2.103615],accel_mss,speed_ms,0,blend_radius_m)
  movel([0.537356, -1.379654, -2.571413, -0.761323, 1.570796, 2.108152],accel_mss,speed_ms,0,blend_radius_m)
  movel([0.542010, -1.377071, -2.573228, -0.762090, 1.570796, 2.112807],accel_mss,speed_ms,0,blend_radius_m)
  movel([0.544261, -1.376252, -2.573801, -0.762335, 1.570796, 2.115058],accel_mss,speed_ms,0,blend_radius_m)
  movel([0.546405, -1.375811, -2.574110, -0.762468, 1.570796, 2.117201],accel_mss,speed_ms,0,blend_radius_m)
  movel([0.548385, -1.375800, -2.574118, -0.762471, 1.570796, 2.119182],accel_mss,speed_ms,0,blend_radius_m)
  movel([0.550163, -1.376263, -2.573794, -0.762332, 1.570796, 2.120959],accel_mss,speed_ms,0,blend_radius_m)
  movel([0.551685, -1.377248, -2.573104, -0.762037, 1.570796, 2.122481],accel_mss,speed_ms,0,blend_radius_m)
  movel([0.552907, -1.378801, -2.572013, -0.761575, 1.570796, 2.123703],accel_mss,speed_ms,0,blend_radius_m)
  movel([0.553764, -1.381691, -2.569974, -0.760724, 1.570796, 2.124560],accel_mss,speed_ms,0,blend_radius_m)
  movel([0.553365, -1.384869, -2.567718, -0.759802, 1.570796, 2.124162],accel_mss,speed_ms,0,blend_radius_m)
  movel([0.551864, -1.388205, -2.565333, -0.758850, 1.570796, 2.122660],accel_mss,speed_ms,0,blend_radius_m)
  movel([0.549416, -1.391581, -2.562905, -0.757903, 1.570796, 2.120212],accel_mss,speed_ms,0,blend_radius_m)
  movel([0.545951, -1.394968, -2.560451, -0.756970, 1.570796, 2.116748],accel_mss,speed_ms,0,blend_radius_m)
  movel([0.542427, -1.397258, -2.558783, -0.756348, 1.570796, 2.113224],accel_mss,speed_ms,0,blend_radius_m)
  movel([0.538901, -1.398590, -2.557808, -0.755990, 1.570796, 2.109697],accel_mss,speed_ms,0,blend_radius_m)
  speed_ms = 0.003
  movel([0.538901, -1.392148, -2.554861, -0.765381, 1.570796, 2.109697],accel_mss,speed_ms,0,blend_radius_m)
  speed_ms = 0.03
  movel([0.538901, -1.367315, -2.542780, -0.802295, 1.570796, 2.109697],accel_mss,speed_ms,0,blend_radius_m)
  #M_RunCode9
  movel([0.645968, -1.263196, -2.608374, -0.840819, 1.570796, 2.216765],accel_mss,speed_ms,0,blend_radius_m)
  #M_RunCode3
  movel([0.645968, -1.289767, -2.621805, -0.800817, 1.570796, 2.216765],accel_mss,speed_ms,0,blend_radius_m)
  speed_ms = 0.003
  movel([0.645968, -1.296710, -2.625093, -0.790586, 1.570796, 2.216765],accel_mss,speed_ms,0,blend_radius_m)
  speed_ms = 0.007
  movel([0.644726, -1.295158, -2.626009, -0.791222, 1.570796, 2.215522],accel_mss,speed_ms,0,blend_radius_m)
  movel([0.644077, -1.293106, -2.627217, -0.792066, 1.570796, 2.214873],accel_mss,speed_ms,0,blend_radius_m)
  movel([0.643766, -1.290803, -2.628565, -0.793021, 1.570796, 2.214562],accel_mss,speed_ms,0,blend_radius_m)
  movel([0.644793, -1.290586, -2.628692, -0.793111, 1.570796, 2.215589],accel_mss,speed_ms,0,blend_radius_m)
  movel([0.645345, -1.291072, -2.628408, -0.792909, 1.570796, 2.216142],accel_mss,speed_ms,0,blend_radius_m)
  movel([0.646043, -1.291573, -2.628115, -0.792701, 1.570796, 2.216839],accel_mss,speed_ms,0,blend_radius_m)
  movel([0.647510, -1.291400, -2.628216, -0.792773, 1.570796, 2.218307],accel_mss,speed_ms,0,blend_radius_m)
  movel([0.649191, -1.290561, -2.628707, -0.793121, 1.570796, 2.219987],accel_mss,speed_ms,0,blend_radius_m)
  movel([0.650832, -1.289421, -2.629371, -0.793597, 1.570796, 2.221629],accel_mss,speed_ms,0,blend_radius_m)
  movel([0.653088, -1.287764, -2.630335, -0.794291, 1.570796, 2.223884],accel_mss,speed_ms,0,blend_radius_m)
  movel([0.652893, -1.284760, -2.632072, -0.795557, 1.570796, 2.223689],accel_mss,speed_ms,0,blend_radius_m)
  movel([0.651858, -1.282725, -2.633242, -0.796422, 1.570796, 2.222655],accel_mss,speed_ms,0,blend_radius_m)
  movel([0.650939, -1.282218, -2.633533, -0.796638, 1.570796, 2.221735],accel_mss,speed_ms,0,blend_radius_m)
  movel([0.649711, -1.282125, -2.633587, -0.796678, 1.570796, 2.220508],accel_mss,speed_ms,0,blend_radius_m)
  movel([0.648143, -1.282504, -2.633369, -0.796516, 1.570796, 2.218939],accel_mss,speed_ms,0,blend_radius_m)
  movel([0.646202, -1.283412, -2.632848, -0.796129, 1.570796, 2.216998],accel_mss,speed_ms,0,blend_radius_m)
  movel([0.647075, -1.281413, -2.633994, -0.796982, 1.570796, 2.217871],accel_mss,speed_ms,0,blend_radius_m)
  movel([0.648052, -1.279711, -2.634966, -0.797712, 1.570796, 2.218848],accel_mss,speed_ms,0,blend_radius_m)
  movel([0.648614, -1.279127, -2.635299, -0.797963, 1.570796, 2.219410],accel_mss,speed_ms,0,blend_radius_m)
  movel([0.649252, -1.278801, -2.635484, -0.798103, 1.570796, 2.220049],accel_mss,speed_ms,0,blend_radius_m)
  movel([0.650801, -1.279188, -2.635264, -0.797937, 1.570796, 2.221597],accel_mss,speed_ms,0,blend_radius_m)
  movel([0.653005, -1.281287, -2.634067, -0.797036, 1.570796, 2.223802],accel_mss,speed_ms,0,blend_radius_m)
  movel([0.654416, -1.284137, -2.632431, -0.795821, 1.570796, 2.225212],accel_mss,speed_ms,0,blend_radius_m)
  movel([0.654640, -1.285774, -2.631487, -0.795128, 1.570796, 2.225436],accel_mss,speed_ms,0,blend_radius_m)
  movel([0.654450, -1.287511, -2.630481, -0.794396, 1.570796, 2.225246],accel_mss,speed_ms,0,blend_radius_m)
  movel([0.653783, -1.289319, -2.629430, -0.793639, 1.570796, 2.224579],accel_mss,speed_ms,0,blend_radius_m)
  movel([0.652561, -1.291170, -2.628351, -0.792868, 1.570796, 2.223357],accel_mss,speed_ms,0,blend_radius_m)
  movel([0.651111, -1.289927, -2.629076, -0.793385, 1.570796, 2.221908],accel_mss,speed_ms,0,blend_radius_m)
  movel([0.648057, -1.297520, -2.624613, -0.790256, 1.570796, 2.218854],accel_mss,speed_ms,0,blend_radius_m)
  movel([0.645968, -1.296710, -2.625093, -0.790586, 1.570796, 2.216765],accel_mss,speed_ms,0,blend_radius_m)
  speed_ms = 0.003
  movel([0.645968, -1.289767, -2.621805, -0.800817, 1.570796, 2.216765],accel_mss,speed_ms,0,blend_radius_m)
  speed_ms = 0.03
  movel([0.645968, -1.263196, -2.608374, -0.840819, 1.570796, 2.216765],accel_mss,speed_ms,0,blend_radius_m)
  #M_RunCode9
  movel([0.625552, -1.207520, -2.637984, -0.866886, 1.570796, 2.196348],accel_mss,speed_ms,0,blend_radius_m)
  #M_RunCode3
  movel([0.625552, -1.234777, -2.652152, -0.825460, 1.570796, 2.196348],accel_mss,speed_ms,0,blend_radius_m)
  speed_ms = 0.003
  movel([0.625552, -1.241929, -2.655627, -0.814833, 1.570796, 2.196348],accel_mss,speed_ms,0,blend_radius_m)
  speed_ms = 0.007
  movel([0.622055, -1.244296, -2.654383, -0.813710, 1.570796, 2.192852],accel_mss,speed_ms,0,blend_radius_m)
  movel([0.618429, -1.246349, -2.653299, -0.812741, 1.570796, 2.189225],accel_mss,speed_ms,0,blend_radius_m)
  movel([0.614714, -1.248050, -2.652397, -0.811942, 1.570796, 2.185511],accel_mss,speed_ms,0,blend_radius_m)
  movel([0.610950, -1.249360, -2.651700, -0.811329, 1.570796, 2.181747],accel_mss,speed_ms,0,blend_radius_m)
  movel([0.607174, -1.250243, -2.651229, -0.810917, 1.570796, 2.177970],accel_mss,speed_ms,0,blend_radius_m)
  movel([0.605296, -1.250294, -2.651202, -0.810893, 1.570796, 2.176092],accel_mss,speed_ms,0,blend_radius_m)
  movel([0.603450, -1.250031, -2.651342, -0.811016, 1.570796, 2.174246],accel_mss,speed_ms,0,blend_radius_m)
  movel([0.601785, -1.249809, -2.651460, -0.811120, 1.570796, 2.172581],accel_mss,speed_ms,0,blend_radius_m)
  movel([0.600456, -1.249976, -2.651372, -0.811042, 1.570796, 2.171252],accel_mss,speed_ms,0,blend_radius_m)
  movel([0.598125, -1.251471, -2.650573, -0.810346, 1.570796, 2.168921],accel_mss,speed_ms,0,blend_radius_m)
  movel([0.595030, -1.253923, -2.649256, -0.809210, 1.570796, 2.165826],accel_mss,speed_ms,0,blend_radius_m)
  movel([0.591820, -1.256516, -2.647856, -0.808017, 1.570796, 2.162617],accel_mss,speed_ms,0,blend_radius_m)
  movel([0.589123, -1.258440, -2.646811, -0.807137, 1.570796, 2.159920],accel_mss,speed_ms,0,blend_radius_m)
  movel([0.583840, -1.261193, -2.645310, -0.805886, 1.570796, 2.154636],accel_mss,speed_ms,0,blend_radius_m)
  movel([0.579153, -1.262895, -2.644377, -0.805117, 1.570796, 2.149949],accel_mss,speed_ms,0,blend_radius_m)
  movel([0.575004, -1.263654, -2.643960, -0.804775, 1.570796, 2.145801],accel_mss,speed_ms,0,blend_radius_m)
  movel([0.571342, -1.263566, -2.644008, -0.804815, 1.570796, 2.142138],accel_mss,speed_ms,0,blend_radius_m)
  movel([0.568117, -1.262730, -2.644467, -0.805191, 1.570796, 2.138913],accel_mss,speed_ms,0,blend_radius_m)
  movel([0.565282, -1.261238, -2.645285, -0.805866, 1.570796, 2.136078],accel_mss,speed_ms,0,blend_radius_m)
  movel([0.562796, -1.259182, -2.646408, -0.806799, 1.570796, 2.133593],accel_mss,speed_ms,0,blend_radius_m)
  movel([0.560619, -1.256653, -2.647781, -0.807954, 1.570796, 2.131415],accel_mss,speed_ms,0,blend_radius_m)
  movel([0.557019, -1.250546, -2.651067, -0.810776, 1.570796, 2.127816],accel_mss,speed_ms,0,blend_radius_m)
  movel([0.554174, -1.243663, -2.654716, -0.814010, 1.570796, 2.124971],accel_mss,speed_ms,0,blend_radius_m)
  movel([0.549511, -1.230699, -2.661438, -0.820252, 1.570796, 2.120307],accel_mss,speed_ms,0,blend_radius_m)
  movel([0.546767, -1.225443, -2.664108, -0.822838, 1.570796, 2.117563],accel_mss,speed_ms,0,blend_radius_m)
  movel([0.542890, -1.219879, -2.666899, -0.825611, 1.570796, 2.113686],accel_mss,speed_ms,0,blend_radius_m)
  movel([0.538028, -1.214344, -2.669641, -0.828404, 1.570796, 2.108824],accel_mss,speed_ms,0,blend_radius_m)
  movel([0.532339, -1.209186, -2.672165, -0.831039, 1.570796, 2.103135],accel_mss,speed_ms,0,blend_radius_m)
  movel([0.525993, -1.204754, -2.674310, -0.833326, 1.570796, 2.096789],accel_mss,speed_ms,0,blend_radius_m)
  movel([0.519181, -1.201391, -2.675923, -0.835075, 1.570796, 2.089978],accel_mss,speed_ms,0,blend_radius_m)
  movel([0.512116, -1.199431, -2.676857, -0.836101, 1.570796, 2.082913],accel_mss,speed_ms,0,blend_radius_m)
  movel([0.508557, -1.199078, -2.677025, -0.836286, 1.570796, 2.079353],accel_mss,speed_ms,0,blend_radius_m)
  movel([0.505021, -1.199191, -2.676971, -0.836227, 1.570796, 2.075817],accel_mss,speed_ms,0,blend_radius_m)
  movel([0.501202, -1.199798, -2.676682, -0.835909, 1.570796, 2.071999],accel_mss,speed_ms,0,blend_radius_m)
  movel([0.496609, -1.200960, -2.676128, -0.835301, 1.570796, 2.067405],accel_mss,speed_ms,0,blend_radius_m)
  movel([0.491506, -1.202720, -2.675287, -0.834382, 1.570796, 2.062302],accel_mss,speed_ms,0,blend_radius_m)
  movel([0.486154, -1.205107, -2.674140, -0.833143, 1.570796, 2.056951],accel_mss,speed_ms,0,blend_radius_m)
  movel([0.480824, -1.208142, -2.672672, -0.831575, 1.570796, 2.051620],accel_mss,speed_ms,0,blend_radius_m)
  movel([0.475782, -1.211850, -2.670865, -0.829674, 1.570796, 2.046578],accel_mss,speed_ms,0,blend_radius_m)
  movel([0.471291, -1.216235, -2.668708, -0.827446, 1.570796, 2.042087],accel_mss,speed_ms,0,blend_radius_m)
  movel([0.469336, -1.218683, -2.667494, -0.826212, 1.570796, 2.040132],accel_mss,speed_ms,0,blend_radius_m)
  movel([0.467617, -1.221306, -2.666186, -0.824897, 1.570796, 2.038413],accel_mss,speed_ms,0,blend_radius_m)
  movel([0.465708, -1.225421, -2.664119, -0.822850, 1.570796, 2.036504],accel_mss,speed_ms,0,blend_radius_m)
  movel([0.465103, -1.228926, -2.662342, -0.821121, 1.570796, 2.035900],accel_mss,speed_ms,0,blend_radius_m)
  movel([0.465645, -1.231885, -2.660831, -0.819673, 1.570796, 2.036441],accel_mss,speed_ms,0,blend_radius_m)
  movel([0.467190, -1.234356, -2.659562, -0.818471, 1.570796, 2.037987],accel_mss,speed_ms,0,blend_radius_m)
  movel([0.469598, -1.236396, -2.658508, -0.817484, 1.570796, 2.040394],accel_mss,speed_ms,0,blend_radius_m)
  movel([0.472726, -1.238064, -2.657644, -0.816681, 1.570796, 2.043522],accel_mss,speed_ms,0,blend_radius_m)
  movel([0.476435, -1.239416, -2.656940, -0.816033, 1.570796, 2.047231],accel_mss,speed_ms,0,blend_radius_m)
  movel([0.480593, -1.240500, -2.656375, -0.815514, 1.570796, 2.051389],accel_mss,speed_ms,0,blend_radius_m)
  movel([0.489718, -1.242066, -2.655555, -0.814768, 1.570796, 2.060515],accel_mss,speed_ms,0,blend_radius_m)
  movel([0.499041, -1.243128, -2.654998, -0.814263, 1.570796, 2.069837],accel_mss,speed_ms,0,blend_radius_m)
  movel([0.507518, -1.244009, -2.654534, -0.813846, 1.570796, 2.078314],accel_mss,speed_ms,0,blend_radius_m)
  movel([0.514107, -1.244994, -2.654015, -0.813380, 1.570796, 2.084903],accel_mss,speed_ms,0,blend_radius_m)
  movel([0.529501, -1.248267, -2.652282, -0.811841, 1.570796, 2.100298],accel_mss,speed_ms,0,blend_radius_m)
  movel([0.537500, -1.250354, -2.651170, -0.810866, 1.570796, 2.108296],accel_mss,speed_ms,0,blend_radius_m)
  movel([0.543400, -1.252488, -2.650027, -0.809874, 1.570796, 2.114196],accel_mss,speed_ms,0,blend_radius_m)
  movel([0.545402, -1.253712, -2.649369, -0.809308, 1.570796, 2.116199],accel_mss,speed_ms,0,blend_radius_m)
  movel([0.547055, -1.255239, -2.648546, -0.808604, 1.570796, 2.117851],accel_mss,speed_ms,0,blend_radius_m)
  movel([0.549358, -1.259078, -2.646464, -0.806846, 1.570796, 2.120154],accel_mss,speed_ms,0,blend_radius_m)
  movel([0.550439, -1.263758, -2.643902, -0.804729, 1.570796, 2.121235],accel_mss,speed_ms,0,blend_radius_m)
  movel([0.550426, -1.269039, -2.640979, -0.802371, 1.570796, 2.121222],accel_mss,speed_ms,0,blend_radius_m)
  movel([0.549452, -1.274685, -2.637816, -0.799888, 1.570796, 2.120249],accel_mss,speed_ms,0,blend_radius_m)
  movel([0.547650, -1.280476, -2.634530, -0.797383, 1.570796, 2.118446],accel_mss,speed_ms,0,blend_radius_m)
  movel([0.545142, -1.286199, -2.631241, -0.794949, 1.570796, 2.115939],accel_mss,speed_ms,0,blend_radius_m)
  movel([0.542048, -1.291646, -2.628072, -0.792670, 1.570796, 2.112844],accel_mss,speed_ms,0,blend_radius_m)
  movel([0.537469, -1.297972, -2.624345, -0.790072, 1.570796, 2.108266],accel_mss,speed_ms,0,blend_radius_m)
  movel([0.535236, -1.300443, -2.622875, -0.789071, 1.570796, 2.106032],accel_mss,speed_ms,0,blend_radius_m)
  movel([0.533018, -1.302518, -2.621634, -0.788237, 1.570796, 2.103815],accel_mss,speed_ms,0,blend_radius_m)
  movel([0.530801, -1.304245, -2.620598, -0.787546, 1.570796, 2.101598],accel_mss,speed_ms,0,blend_radius_m)
  movel([0.528569, -1.305669, -2.619740, -0.786980, 1.570796, 2.099365],accel_mss,speed_ms,0,blend_radius_m)
  movel([0.524002, -1.307779, -2.618464, -0.786146, 1.570796, 2.094798],accel_mss,speed_ms,0,blend_radius_m)
  movel([0.519208, -1.309197, -2.617603, -0.785589, 1.570796, 2.090004],accel_mss,speed_ms,0,blend_radius_m)
  movel([0.514074, -1.310271, -2.616950, -0.785168, 1.570796, 2.084870],accel_mss,speed_ms,0,blend_radius_m)
  movel([0.502416, -1.312726, -2.615450, -0.784213, 1.570796, 2.073212],accel_mss,speed_ms,0,blend_radius_m)
  movel([0.501805, -1.312910, -2.615337, -0.784142, 1.570796, 2.072602],accel_mss,speed_ms,0,blend_radius_m)
  movel([0.501991, -1.313037, -2.615259, -0.784093, 1.570796, 2.072788],accel_mss,speed_ms,0,blend_radius_m)
  movel([0.504325, -1.313158, -2.615185, -0.784046, 1.570796, 2.075121],accel_mss,speed_ms,0,blend_radius_m)
  movel([0.513941, -1.313094, -2.615224, -0.784071, 1.570796, 2.084738],accel_mss,speed_ms,0,blend_radius_m)
  movel([0.529835, -1.313150, -2.615190, -0.784049, 1.570796, 2.100631],accel_mss,speed_ms,0,blend_radius_m)
  movel([0.520283, -1.317184, -2.612706, -0.782499, 1.570796, 2.091080],accel_mss,speed_ms,0,blend_radius_m)
  movel([0.509692, -1.321219, -2.610200, -0.780970, 1.570796, 2.080488],accel_mss,speed_ms,0,blend_radius_m)
  movel([0.498438, -1.325183, -2.607716, -0.779489, 1.570796, 2.069234],accel_mss,speed_ms,0,blend_radius_m)
  movel([0.486893, -1.329003, -2.605303, -0.778082, 1.570796, 2.057689],accel_mss,speed_ms,0,blend_radius_m)
  movel([0.464414, -1.335840, -2.600935, -0.775613, 1.570796, 2.035210],accel_mss,speed_ms,0,blend_radius_m)
  movel([0.454207, -1.338650, -2.599122, -0.774617, 1.570796, 2.025004],accel_mss,speed_ms,0,blend_radius_m)
  movel([0.445174, -1.340897, -2.597664, -0.773828, 1.570796, 2.015971],accel_mss,speed_ms,0,blend_radius_m)
  movel([0.432414, -1.348751, -2.592514, -0.771124, 1.570796, 2.003210],accel_mss,speed_ms,0,blend_radius_m)
  movel([0.419549, -1.357340, -2.586784, -0.768265, 1.570796, 1.990346],accel_mss,speed_ms,0,blend_radius_m)
  movel([0.393955, -1.375427, -2.574378, -0.762583, 1.570796, 1.964752],accel_mss,speed_ms,0,blend_radius_m)
  movel([0.381401, -1.384334, -2.568099, -0.759956, 1.570796, 1.952197],accel_mss,speed_ms,0,blend_radius_m)
  movel([0.369096, -1.392783, -2.562036, -0.757570, 1.570796, 1.939892],accel_mss,speed_ms,0,blend_radius_m)
  movel([0.357076, -1.400519, -2.556393, -0.755476, 1.570796, 1.927872],accel_mss,speed_ms,0,blend_radius_m)
  movel([0.345373, -1.407305, -2.551372, -0.753712, 1.570796, 1.916169],accel_mss,speed_ms,0,blend_radius_m)
  movel([0.340839, -1.409583, -2.549671, -0.753135, 1.570796, 1.911635],accel_mss,speed_ms,0,blend_radius_m)
  movel([0.336536, -1.411411, -2.548301, -0.752677, 1.570796, 1.907333],accel_mss,speed_ms,0,blend_radius_m)
  movel([0.332488, -1.412794, -2.547260, -0.752334, 1.570796, 1.903284],accel_mss,speed_ms,0,blend_radius_m)
  movel([0.328710, -1.413736, -2.546550, -0.752103, 1.570796, 1.899506],accel_mss,speed_ms,0,blend_radius_m)
  movel([0.325228, -1.414239, -2.546170, -0.751979, 1.570796, 1.896024],accel_mss,speed_ms,0,blend_radius_m)
  movel([0.322064, -1.414307, -2.546119, -0.751963, 1.570796, 1.892861],accel_mss,speed_ms,0,blend_radius_m)
  movel([0.319239, -1.413938, -2.546398, -0.752053, 1.570796, 1.890036],accel_mss,speed_ms,0,blend_radius_m)
  movel([0.316779, -1.413136, -2.547003, -0.752250, 1.570796, 1.887576],accel_mss,speed_ms,0,blend_radius_m)
  movel([0.314710, -1.411894, -2.547938, -0.752557, 1.570796, 1.885507],accel_mss,speed_ms,0,blend_radius_m)
  movel([0.313060, -1.410214, -2.549198, -0.752976, 1.570796, 1.883856],accel_mss,speed_ms,0,blend_radius_m)
  movel([0.311851, -1.408094, -2.550784, -0.753511, 1.570796, 1.882648],accel_mss,speed_ms,0,blend_radius_m)
  movel([0.311120, -1.405524, -2.552696, -0.754168, 1.570796, 1.881917],accel_mss,speed_ms,0,blend_radius_m)
  movel([0.310896, -1.402502, -2.554933, -0.754954, 1.570796, 1.881693],accel_mss,speed_ms,0,blend_radius_m)
  movel([0.311213, -1.399021, -2.557493, -0.755875, 1.570796, 1.882009],accel_mss,speed_ms,0,blend_radius_m)
  movel([0.312103, -1.395073, -2.560375, -0.756941, 1.570796, 1.882900],accel_mss,speed_ms,0,blend_radius_m)
  movel([0.313607, -1.390651, -2.563575, -0.758162, 1.570796, 1.884403],accel_mss,speed_ms,0,blend_radius_m)
  movel([0.317142, -1.391966, -2.562627, -0.757796, 1.570796, 1.887939],accel_mss,speed_ms,0,blend_radius_m)
  movel([0.318943, -1.392493, -2.562245, -0.757650, 1.570796, 1.889739],accel_mss,speed_ms,0,blend_radius_m)
  movel([0.320933, -1.392540, -2.562211, -0.757637, 1.570796, 1.891729],accel_mss,speed_ms,0,blend_radius_m)
  movel([0.322664, -1.392046, -2.562569, -0.757774, 1.570796, 1.893460],accel_mss,speed_ms,0,blend_radius_m)
  movel([0.324819, -1.391028, -2.563304, -0.758057, 1.570796, 1.895616],accel_mss,speed_ms,0,blend_radius_m)
  movel([0.330186, -1.387662, -2.565723, -0.759004, 1.570796, 1.900983],accel_mss,speed_ms,0,blend_radius_m)
  movel([0.336585, -1.382956, -2.569078, -0.760356, 1.570796, 1.907381],accel_mss,speed_ms,0,blend_radius_m)
  movel([0.343564, -1.377417, -2.572985, -0.761987, 1.570796, 1.914360],accel_mss,speed_ms,0,blend_radius_m)
  movel([0.357335, -1.365936, -2.580945, -0.765507, 1.570796, 1.928131],accel_mss,speed_ms,0,blend_radius_m)
  movel([0.367417, -1.357545, -2.586646, -0.768199, 1.570796, 1.938214],accel_mss,speed_ms,0,blend_radius_m)
  movel([0.376504, -1.350810, -2.591150, -0.770430, 1.570796, 1.947300],accel_mss,speed_ms,0,blend_radius_m)
  movel([0.385701, -1.344042, -2.595612, -0.772735, 1.570796, 1.956498],accel_mss,speed_ms,0,blend_radius_m)
  movel([0.367254, -1.347443, -2.593377, -0.771569, 1.570796, 1.938050],accel_mss,speed_ms,0,blend_radius_m)
  movel([0.357739, -1.348863, -2.592440, -0.771086, 1.570796, 1.928535],accel_mss,speed_ms,0,blend_radius_m)
  movel([0.348701, -1.349461, -2.592044, -0.770884, 1.570796, 1.919497],accel_mss,speed_ms,0,blend_radius_m)
  movel([0.344513, -1.349300, -2.592151, -0.770939, 1.570796, 1.915310],accel_mss,speed_ms,0,blend_radius_m)
  movel([0.340630, -1.348747, -2.592516, -0.771126, 1.570796, 1.911427],accel_mss,speed_ms,0,blend_radius_m)
  movel([0.337108, -1.347741, -2.593181, -0.771467, 1.570796, 1.907905],accel_mss,speed_ms,0,blend_radius_m)
  movel([0.334013, -1.346214, -2.594186, -0.771988, 1.570796, 1.904809],accel_mss,speed_ms,0,blend_radius_m)
  movel([0.331406, -1.344096, -2.595577, -0.772716, 1.570796, 1.902202],accel_mss,speed_ms,0,blend_radius_m)
  movel([0.329346, -1.341321, -2.597388, -0.773680, 1.570796, 1.900142],accel_mss,speed_ms,0,blend_radius_m)
  movel([0.327906, -1.337812, -2.599664, -0.774913, 1.570796, 1.898703],accel_mss,speed_ms,0,blend_radius_m)
  movel([0.327152, -1.333488, -2.602445, -0.776455, 1.570796, 1.897948],accel_mss,speed_ms,0,blend_radius_m)
  movel([0.327355, -1.327896, -2.606005, -0.778488, 1.570796, 1.898151],accel_mss,speed_ms,0,blend_radius_m)
  movel([0.328755, -1.321784, -2.609847, -0.780758, 1.570796, 1.899551],accel_mss,speed_ms,0,blend_radius_m)
  movel([0.331266, -1.315338, -2.613845, -0.783206, 1.570796, 1.902062],accel_mss,speed_ms,0,blend_radius_m)
  movel([0.334788, -1.308757, -2.617871, -0.785761, 1.570796, 1.905584],accel_mss,speed_ms,0,blend_radius_m)
  movel([0.339224, -1.302255, -2.621792, -0.788342, 1.570796, 1.910020],accel_mss,speed_ms,0,blend_radius_m)
  movel([0.344458, -1.296055, -2.625480, -0.790854, 1.570796, 1.915255],accel_mss,speed_ms,0,blend_radius_m)
  movel([0.350374, -1.290391, -2.628806, -0.793192, 1.570796, 1.921170],accel_mss,speed_ms,0,blend_radius_m)
  movel([0.356842, -1.285507, -2.631641, -0.795241, 1.570796, 1.927638],accel_mss,speed_ms,0,blend_radius_m)
  movel([0.360543, -1.283617, -2.632730, -0.796042, 1.570796, 1.931339],accel_mss,speed_ms,0,blend_radius_m)
  movel([0.364662, -1.282307, -2.633482, -0.796600, 1.570796, 1.935458],accel_mss,speed_ms,0,blend_radius_m)
  movel([0.367875, -1.282068, -2.633619, -0.796702, 1.570796, 1.938672],accel_mss,speed_ms,0,blend_radius_m)
  movel([0.368725, -1.282503, -2.633370, -0.796516, 1.570796, 1.939521],accel_mss,speed_ms,0,blend_radius_m)
  movel([0.368853, -1.283383, -2.632864, -0.796141, 1.570796, 1.939650],accel_mss,speed_ms,0,blend_radius_m)
  movel([0.365604, -1.284361, -2.632302, -0.795726, 1.570796, 1.936401],accel_mss,speed_ms,0,blend_radius_m)
  movel([0.362817, -1.285527, -2.631629, -0.795233, 1.570796, 1.933614],accel_mss,speed_ms,0,blend_radius_m)
  movel([0.360485, -1.286847, -2.630866, -0.794676, 1.570796, 1.931281],accel_mss,speed_ms,0,blend_radius_m)
  movel([0.358588, -1.288287, -2.630031, -0.794071, 1.570796, 1.929384],accel_mss,speed_ms,0,blend_radius_m)
  movel([0.357110, -1.289820, -2.629139, -0.793430, 1.570796, 1.927906],accel_mss,speed_ms,0,blend_radius_m)
  movel([0.356041, -1.291411, -2.628210, -0.792768, 1.570796, 1.926837],accel_mss,speed_ms,0,blend_radius_m)
  movel([0.355357, -1.293034, -2.627259, -0.792096, 1.570796, 1.926154],accel_mss,speed_ms,0,blend_radius_m)
  movel([0.355048, -1.294659, -2.626303, -0.791426, 1.570796, 1.925845],accel_mss,speed_ms,0,blend_radius_m)
  movel([0.355479, -1.297808, -2.624442, -0.790139, 1.570796, 1.926275],accel_mss,speed_ms,0,blend_radius_m)
  movel([0.357193, -1.300636, -2.622760, -0.788993, 1.570796, 1.927989],accel_mss,speed_ms,0,blend_radius_m)
  movel([0.360059, -1.302940, -2.621381, -0.788068, 1.570796, 1.930855],accel_mss,speed_ms,0,blend_radius_m)
  movel([0.363953, -1.304506, -2.620441, -0.787442, 1.570796, 1.934749],accel_mss,speed_ms,0,blend_radius_m)
  movel([0.366667, -1.304911, -2.620197, -0.787281, 1.570796, 1.937464],accel_mss,speed_ms,0,blend_radius_m)
  movel([0.370152, -1.304976, -2.620157, -0.787255, 1.570796, 1.940949],accel_mss,speed_ms,0,blend_radius_m)
  movel([0.379029, -1.304255, -2.620592, -0.787542, 1.570796, 1.949825],accel_mss,speed_ms,0,blend_radius_m)
  movel([0.389764, -1.302670, -2.621544, -0.788176, 1.570796, 1.960560],accel_mss,speed_ms,0,blend_radius_m)
  movel([0.401550, -1.300532, -2.622822, -0.789035, 1.570796, 1.972346],accel_mss,speed_ms,0,blend_radius_m)
  movel([0.424998, -1.295719, -2.625678, -0.790992, 1.570796, 1.995795],accel_mss,speed_ms,0,blend_radius_m)
  movel([0.442799, -1.291795, -2.627986, -0.792609, 1.570796, 2.013595],accel_mss,speed_ms,0,blend_radius_m)
  movel([0.451768, -1.289823, -2.629137, -0.793429, 1.570796, 2.022565],accel_mss,speed_ms,0,blend_radius_m)
  movel([0.456636, -1.288609, -2.629844, -0.793936, 1.570796, 2.027432],accel_mss,speed_ms,0,blend_radius_m)
  movel([0.460382, -1.287357, -2.630571, -0.794461, 1.570796, 2.031178],accel_mss,speed_ms,0,blend_radius_m)
  movel([0.461423, -1.286797, -2.630895, -0.794697, 1.570796, 2.032219],accel_mss,speed_ms,0,blend_radius_m)
  movel([0.461864, -1.286278, -2.631195, -0.794916, 1.570796, 2.032661],accel_mss,speed_ms,0,blend_radius_m)
  movel([0.461437, -1.285089, -2.631882, -0.795418, 1.570796, 2.032234],accel_mss,speed_ms,0,blend_radius_m)
  movel([0.458790, -1.282637, -2.633293, -0.796459, 1.570796, 2.029586],accel_mss,speed_ms,0,blend_radius_m)
  movel([0.455344, -1.280813, -2.634337, -0.797239, 1.570796, 2.026140],accel_mss,speed_ms,0,blend_radius_m)
  movel([0.447553, -1.277352, -2.636307, -0.798729, 1.570796, 2.018350],accel_mss,speed_ms,0,blend_radius_m)
  movel([0.443954, -1.274842, -2.637727, -0.799820, 1.570796, 2.014750],accel_mss,speed_ms,0,blend_radius_m)
  movel([0.441047, -1.271211, -2.639767, -0.801411, 1.570796, 2.011844],accel_mss,speed_ms,0,blend_radius_m)
  movel([0.439972, -1.268831, -2.641095, -0.802463, 1.570796, 2.010768],accel_mss,speed_ms,0,blend_radius_m)
  movel([0.439212, -1.265988, -2.642672, -0.803729, 1.570796, 2.010009],accel_mss,speed_ms,0,blend_radius_m)
  movel([0.438817, -1.262623, -2.644526, -0.805240, 1.570796, 2.009614],accel_mss,speed_ms,0,blend_radius_m)
  movel([0.438842, -1.258671, -2.646686, -0.807032, 1.570796, 2.009638],accel_mss,speed_ms,0,blend_radius_m)
  movel([0.439690, -1.253131, -2.649682, -0.809576, 1.570796, 2.010486],accel_mss,speed_ms,0,blend_radius_m)
  movel([0.441519, -1.247582, -2.652646, -0.812162, 1.570796, 2.012315],accel_mss,speed_ms,0,blend_radius_m)
  movel([0.444219, -1.242044, -2.655567, -0.814779, 1.570796, 2.015015],accel_mss,speed_ms,0,blend_radius_m)
  movel([0.447687, -1.236534, -2.658437, -0.817418, 1.570796, 2.018484],accel_mss,speed_ms,0,blend_radius_m)
  movel([0.451801, -1.231077, -2.661245, -0.820067, 1.570796, 2.022598],accel_mss,speed_ms,0,blend_radius_m)
  movel([0.456447, -1.225700, -2.663978, -0.822711, 1.570796, 2.027243],accel_mss,speed_ms,0,blend_radius_m)
  movel([0.461503, -1.220424, -2.666627, -0.825338, 1.570796, 2.032299],accel_mss,speed_ms,0,blend_radius_m)
  movel([0.466849, -1.215279, -2.669180, -0.827930, 1.570796, 2.037646],accel_mss,speed_ms,0,blend_radius_m)
  movel([0.477396, -1.206212, -2.673606, -0.832571, 1.570796, 2.048192],accel_mss,speed_ms,0,blend_radius_m)
  movel([0.487066, -1.199131, -2.676999, -0.836258, 1.570796, 2.057862],accel_mss,speed_ms,0,blend_radius_m)
  movel([0.495379, -1.193942, -2.679451, -0.838996, 1.570796, 2.066176],accel_mss,speed_ms,0,blend_radius_m)
  movel([0.501871, -1.190519, -2.681052, -0.840818, 1.570796, 2.072668],accel_mss,speed_ms,0,blend_radius_m)
  movel([0.511450, -1.186590, -2.682875, -0.842924, 1.570796, 2.082246],accel_mss,speed_ms,0,blend_radius_m)
  movel([0.520613, -1.184083, -2.684029, -0.844277, 1.570796, 2.091410],accel_mss,speed_ms,0,blend_radius_m)
  movel([0.529237, -1.182967, -2.684540, -0.844881, 1.570796, 2.100033],accel_mss,speed_ms,0,blend_radius_m)
  movel([0.537203, -1.183208, -2.684430, -0.844751, 1.570796, 2.108000],accel_mss,speed_ms,0,blend_radius_m)
  movel([0.544404, -1.184751, -2.683722, -0.843916, 1.570796, 2.115201],accel_mss,speed_ms,0,blend_radius_m)
  movel([0.550735, -1.187532, -2.682439, -0.842418, 1.570796, 2.121531],accel_mss,speed_ms,0,blend_radius_m)
  movel([0.556113, -1.191471, -2.680608, -0.840309, 1.570796, 2.126909],accel_mss,speed_ms,0,blend_radius_m)
  movel([0.560458, -1.196483, -2.678254, -0.837652, 1.570796, 2.131255],accel_mss,speed_ms,0,blend_radius_m)
  movel([0.563420, -1.201840, -2.675708, -0.834841, 1.570796, 2.134216],accel_mss,speed_ms,0,blend_radius_m)
  movel([0.565757, -1.207618, -2.672926, -0.831845, 1.570796, 2.136553],accel_mss,speed_ms,0,blend_radius_m)
  movel([0.567934, -1.213357, -2.670126, -0.828906, 1.570796, 2.138730],accel_mss,speed_ms,0,blend_radius_m)
  movel([0.570419, -1.218631, -2.667520, -0.826238, 1.570796, 2.141215],accel_mss,speed_ms,0,blend_radius_m)
  movel([0.573657, -1.223026, -2.665325, -0.824039, 1.570796, 2.144453],accel_mss,speed_ms,0,blend_radius_m)
  movel([0.575701, -1.224769, -2.664448, -0.823173, 1.570796, 2.146497],accel_mss,speed_ms,0,blend_radius_m)
  movel([0.578105, -1.226144, -2.663754, -0.822492, 1.570796, 2.148902],accel_mss,speed_ms,0,blend_radius_m)
  movel([0.580922, -1.227105, -2.663267, -0.822017, 1.570796, 2.151718],accel_mss,speed_ms,0,blend_radius_m)
  movel([0.584212, -1.227604, -2.663014, -0.821771, 1.570796, 2.155008],accel_mss,speed_ms,0,blend_radius_m)
  movel([0.588036, -1.227587, -2.663022, -0.821779, 1.570796, 2.158832],accel_mss,speed_ms,0,blend_radius_m)
  movel([0.592450, -1.227015, -2.663312, -0.822061, 1.570796, 2.163247],accel_mss,speed_ms,0,blend_radius_m)
  movel([0.596503, -1.225902, -2.663876, -0.822611, 1.570796, 2.167299],accel_mss,speed_ms,0,blend_radius_m)
  movel([0.600105, -1.224204, -2.664732, -0.823453, 1.570796, 2.170902],accel_mss,speed_ms,0,blend_radius_m)
  movel([0.603248, -1.222025, -2.665826, -0.824537, 1.570796, 2.174045],accel_mss,speed_ms,0,blend_radius_m)
  movel([0.605926, -1.219476, -2.667100, -0.825814, 1.570796, 2.176722],accel_mss,speed_ms,0,blend_radius_m)
  movel([0.608121, -1.216664, -2.668496, -0.827230, 1.570796, 2.178918],accel_mss,speed_ms,0,blend_radius_m)
  movel([0.609818, -1.213704, -2.669955, -0.828730, 1.570796, 2.180614],accel_mss,speed_ms,0,blend_radius_m)
  movel([0.611005, -1.210710, -2.671422, -0.830257, 1.570796, 2.181801],accel_mss,speed_ms,0,blend_radius_m)
  movel([0.611653, -1.207806, -2.672835, -0.831748, 1.570796, 2.182449],accel_mss,speed_ms,0,blend_radius_m)
  movel([0.611748, -1.205110, -2.674138, -0.833141, 1.570796, 2.182544],accel_mss,speed_ms,0,blend_radius_m)
  movel([0.611269, -1.202750, -2.675272, -0.834367, 1.570796, 2.182066],accel_mss,speed_ms,0,blend_radius_m)
  movel([0.610196, -1.200855, -2.676179, -0.835356, 1.570796, 2.180992],accel_mss,speed_ms,0,blend_radius_m)
  movel([0.608512, -1.199549, -2.676801, -0.836039, 1.570796, 2.179309],accel_mss,speed_ms,0,blend_radius_m)
  movel([0.606200, -1.198961, -2.677080, -0.836347, 1.570796, 2.176997],accel_mss,speed_ms,0,blend_radius_m)
  movel([0.603247, -1.199219, -2.676958, -0.836212, 1.570796, 2.174043],accel_mss,speed_ms,0,blend_radius_m)
  movel([0.599649, -1.200441, -2.676376, -0.835572, 1.570796, 2.170445],accel_mss,speed_ms,0,blend_radius_m)
  movel([0.595400, -1.202746, -2.675274, -0.834369, 1.570796, 2.166196],accel_mss,speed_ms,0,blend_radius_m)
  movel([0.597575, -1.203321, -2.674998, -0.834069, 1.570796, 2.168372],accel_mss,speed_ms,0,blend_radius_m)
  movel([0.599068, -1.204332, -2.674513, -0.833544, 1.570796, 2.169865],accel_mss,speed_ms,0,blend_radius_m)
  movel([0.599872, -1.205697, -2.673855, -0.832837, 1.570796, 2.170669],accel_mss,speed_ms,0,blend_radius_m)
  movel([0.599986, -1.207348, -2.673057, -0.831984, 1.570796, 2.170782],accel_mss,speed_ms,0,blend_radius_m)
  movel([0.599404, -1.209217, -2.672150, -0.831023, 1.570796, 2.170201],accel_mss,speed_ms,0,blend_radius_m)
  movel([0.598129, -1.211229, -2.671169, -0.829992, 1.570796, 2.168925],accel_mss,speed_ms,0,blend_radius_m)
  movel([0.596156, -1.213321, -2.670143, -0.828924, 1.570796, 2.166953],accel_mss,speed_ms,0,blend_radius_m)
  movel([0.593485, -1.215429, -2.669106, -0.827854, 1.570796, 2.164281],accel_mss,speed_ms,0,blend_radius_m)
  movel([0.588659, -1.218209, -2.667730, -0.826450, 1.570796, 2.159455],accel_mss,speed_ms,0,blend_radius_m)
  movel([0.584354, -1.219614, -2.667031, -0.825744, 1.570796, 2.155151],accel_mss,speed_ms,0,blend_radius_m)
  movel([0.580578, -1.219788, -2.666944, -0.825657, 1.570796, 2.151375],accel_mss,speed_ms,0,blend_radius_m)
  movel([0.577353, -1.218874, -2.667399, -0.826116, 1.570796, 2.148149],accel_mss,speed_ms,0,blend_radius_m)
  movel([0.574703, -1.216990, -2.668334, -0.827065, 1.570796, 2.145499],accel_mss,speed_ms,0,blend_radius_m)
  movel([0.572660, -1.214266, -2.669679, -0.828444, 1.570796, 2.143456],accel_mss,speed_ms,0,blend_radius_m)
  movel([0.571258, -1.210820, -2.671368, -0.830201, 1.570796, 2.142054],accel_mss,speed_ms,0,blend_radius_m)
  movel([0.570539, -1.206770, -2.673337, -0.832282, 1.570796, 2.141335],accel_mss,speed_ms,0,blend_radius_m)
  movel([0.570543, -1.202237, -2.675518, -0.834634, 1.570796, 2.141339],accel_mss,speed_ms,0,blend_radius_m)
  movel([0.571323, -1.197342, -2.677848, -0.837199, 1.570796, 2.142119],accel_mss,speed_ms,0,blend_radius_m)
  movel([0.572919, -1.192208, -2.680264, -0.839917, 1.570796, 2.143715],accel_mss,speed_ms,0,blend_radius_m)
  movel([0.575384, -1.186970, -2.682699, -0.842720, 1.570796, 2.146180],accel_mss,speed_ms,0,blend_radius_m)
  movel([0.578760, -1.181762, -2.685091, -0.845535, 1.570796, 2.149557],accel_mss,speed_ms,0,blend_radius_m)
  movel([0.583096, -1.176730, -2.687375, -0.848284, 1.570796, 2.153893],accel_mss,speed_ms,0,blend_radius_m)
  movel([0.588428, -1.172029, -2.689485, -0.850875, 1.570796, 2.159224],accel_mss,speed_ms,0,blend_radius_m)
  movel([0.594789, -1.167827, -2.691351, -0.853212, 1.570796, 2.165585],accel_mss,speed_ms,0,blend_radius_m)
  movel([0.599497, -1.165367, -2.692434, -0.854587, 1.570796, 2.170293],accel_mss,speed_ms,0,blend_radius_m)
  movel([0.604158, -1.163345, -2.693321, -0.855723, 1.570796, 2.174954],accel_mss,speed_ms,0,blend_radius_m)
  movel([0.608729, -1.161764, -2.694011, -0.856614, 1.570796, 2.179526],accel_mss,speed_ms,0,blend_radius_m)
  movel([0.613176, -1.160631, -2.694504, -0.857254, 1.570796, 2.183972],accel_mss,speed_ms,0,blend_radius_m)
  movel([0.617448, -1.159958, -2.694796, -0.857635, 1.570796, 2.188245],accel_mss,speed_ms,0,blend_radius_m)
  movel([0.621511, -1.159747, -2.694888, -0.857755, 1.570796, 2.192307],accel_mss,speed_ms,0,blend_radius_m)
  movel([0.625325, -1.160000, -2.694778, -0.857611, 1.570796, 2.196121],accel_mss,speed_ms,0,blend_radius_m)
  movel([0.628853, -1.160715, -2.694467, -0.857206, 1.570796, 2.199650],accel_mss,speed_ms,0,blend_radius_m)
  movel([0.632051, -1.161899, -2.693952, -0.856538, 1.570796, 2.202847],accel_mss,speed_ms,0,blend_radius_m)
  movel([0.634891, -1.163547, -2.693232, -0.855609, 1.570796, 2.205687],accel_mss,speed_ms,0,blend_radius_m)
  movel([0.637332, -1.165654, -2.692308, -0.854427, 1.570796, 2.208128],accel_mss,speed_ms,0,blend_radius_m)
  movel([0.639342, -1.168215, -2.691179, -0.852995, 1.570796, 2.210138],accel_mss,speed_ms,0,blend_radius_m)
  movel([0.640896, -1.171221, -2.689845, -0.851323, 1.570796, 2.211693],accel_mss,speed_ms,0,blend_radius_m)
  movel([0.641954, -1.174670, -2.688303, -0.849417, 1.570796, 2.212750],accel_mss,speed_ms,0,blend_radius_m)
  movel([0.642493, -1.178549, -2.686553, -0.847287, 1.570796, 2.213290],accel_mss,speed_ms,0,blend_radius_m)
  movel([0.642488, -1.182847, -2.684595, -0.844947, 1.570796, 2.213285],accel_mss,speed_ms,0,blend_radius_m)
  movel([0.641414, -1.187531, -2.682440, -0.842418, 1.570796, 2.212211],accel_mss,speed_ms,0,blend_radius_m)
  movel([0.639387, -1.192810, -2.679982, -0.839597, 1.570796, 2.210184],accel_mss,speed_ms,0,blend_radius_m)
  movel([0.637426, -1.197366, -2.677837, -0.837186, 1.570796, 2.208223],accel_mss,speed_ms,0,blend_radius_m)
  movel([0.636519, -1.199923, -2.676623, -0.835843, 1.570796, 2.207316],accel_mss,speed_ms,0,blend_radius_m)
  movel([0.637332, -1.201268, -2.675981, -0.835140, 1.570796, 2.208128],accel_mss,speed_ms,0,blend_radius_m)
  movel([0.639265, -1.202921, -2.675190, -0.834278, 1.570796, 2.210061],accel_mss,speed_ms,0,blend_radius_m)
  movel([0.641389, -1.204745, -2.674314, -0.833330, 1.570796, 2.212185],accel_mss,speed_ms,0,blend_radius_m)
  movel([0.642801, -1.206581, -2.673428, -0.832380, 1.570796, 2.213598],accel_mss,speed_ms,0,blend_radius_m)
  movel([0.643727, -1.209704, -2.671912, -0.830772, 1.570796, 2.214523],accel_mss,speed_ms,0,blend_radius_m)
  movel([0.644001, -1.212988, -2.670307, -0.829094, 1.570796, 2.214797],accel_mss,speed_ms,0,blend_radius_m)
  movel([0.643673, -1.216381, -2.668635, -0.827372, 1.570796, 2.214469],accel_mss,speed_ms,0,blend_radius_m)
  movel([0.642802, -1.219834, -2.666921, -0.825634, 1.570796, 2.213598],accel_mss,speed_ms,0,blend_radius_m)
  movel([0.641431, -1.223301, -2.665186, -0.823902, 1.570796, 2.212227],accel_mss,speed_ms,0,blend_radius_m)
  movel([0.639617, -1.226734, -2.663455, -0.822200, 1.570796, 2.210413],accel_mss,speed_ms,0,blend_radius_m)
  movel([0.637410, -1.230090, -2.661749, -0.820550, 1.570796, 2.208206],accel_mss,speed_ms,0,blend_radius_m)
  movel([0.634852, -1.233328, -2.660091, -0.818970, 1.570796, 2.205648],accel_mss,speed_ms,0,blend_radius_m)
  movel([0.631992, -1.236408, -2.658502, -0.817479, 1.570796, 2.202788],accel_mss,speed_ms,0,blend_radius_m)
  movel([0.628880, -1.239287, -2.657007, -0.816095, 1.570796, 2.199676],accel_mss,speed_ms,0,blend_radius_m)
  movel([0.625552, -1.241929, -2.655627, -0.814833, 1.570796, 2.196348],accel_mss,speed_ms,0,blend_radius_m)
  speed_ms = 0.003
  movel([0.625552, -1.234777, -2.652152, -0.825460, 1.570796, 2.196348],accel_mss,speed_ms,0,blend_radius_m)
  speed_ms = 0.03
  movel([0.625552, -1.207520, -2.637984, -0.866886, 1.570796, 2.196348],accel_mss,speed_ms,0,blend_radius_m)
  #M_RunCode9
  movel([0.646760, -1.207578, -2.637954, -0.866856, 1.570796, 2.217556],accel_mss,speed_ms,0,blend_radius_m)
  #M_RunCode3
  movel([0.646760, -1.234835, -2.652122, -0.825432, 1.570796, 2.217556],accel_mss,speed_ms,0,blend_radius_m)
  speed_ms = 0.003
  movel([0.646760, -1.241987, -2.655596, -0.814805, 1.570796, 2.217556],accel_mss,speed_ms,0,blend_radius_m)
  speed_ms = 0.007
  movel([0.648229, -1.239143, -2.657082, -0.816164, 1.570796, 2.219025],accel_mss,speed_ms,0,blend_radius_m)
  movel([0.651947, -1.233399, -2.660054, -0.818935, 1.570796, 2.222744],accel_mss,speed_ms,0,blend_radius_m)
  movel([0.655349, -1.227741, -2.662945, -0.821704, 1.570796, 2.226145],accel_mss,speed_ms,0,blend_radius_m)
  movel([0.656410, -1.225004, -2.664329, -0.823056, 1.570796, 2.227206],accel_mss,speed_ms,0,blend_radius_m)
  movel([0.656763, -1.222366, -2.665655, -0.824367, 1.570796, 2.227559],accel_mss,speed_ms,0,blend_radius_m)
  movel([0.657167, -1.224002, -2.664834, -0.823553, 1.570796, 2.227963],accel_mss,speed_ms,0,blend_radius_m)
  movel([0.657185, -1.227314, -2.663161, -0.821914, 1.570796, 2.227982],accel_mss,speed_ms,0,blend_radius_m)
  movel([0.656357, -1.230634, -2.661471, -0.820284, 1.570796, 2.227153],accel_mss,speed_ms,0,blend_radius_m)
  movel([0.654948, -1.233961, -2.659765, -0.818663, 1.570796, 2.225744],accel_mss,speed_ms,0,blend_radius_m)
  movel([0.653223, -1.237290, -2.658045, -0.817054, 1.570796, 2.224020],accel_mss,speed_ms,0,blend_radius_m)
  movel([0.649856, -1.243951, -2.654565, -0.813873, 1.570796, 2.220653],accel_mss,speed_ms,0,blend_radius_m)
  movel([0.648723, -1.247278, -2.652807, -0.812304, 1.570796, 2.219520],accel_mss,speed_ms,0,blend_radius_m)
  movel([0.648292, -1.250602, -2.651037, -0.810750, 1.570796, 2.219088],accel_mss,speed_ms,0,blend_radius_m)
  movel([0.648584, -1.254052, -2.649186, -0.809151, 1.570796, 2.219380],accel_mss,speed_ms,0,blend_radius_m)
  movel([0.648935, -1.255797, -2.648245, -0.808347, 1.570796, 2.219731],accel_mss,speed_ms,0,blend_radius_m)
  movel([0.649415, -1.256641, -2.647788, -0.807960, 1.570796, 2.220211],accel_mss,speed_ms,0,blend_radius_m)
  movel([0.651300, -1.256077, -2.648093, -0.808219, 1.570796, 2.222097],accel_mss,speed_ms,0,blend_radius_m)
  movel([0.652835, -1.255692, -2.648301, -0.808395, 1.570796, 2.223631],accel_mss,speed_ms,0,blend_radius_m)
  movel([0.654320, -1.255606, -2.648348, -0.808435, 1.570796, 2.225117],accel_mss,speed_ms,0,blend_radius_m)
  movel([0.656913, -1.256158, -2.648049, -0.808181, 1.570796, 2.227710],accel_mss,speed_ms,0,blend_radius_m)
  movel([0.658565, -1.257046, -2.647568, -0.807774, 1.570796, 2.229362],accel_mss,speed_ms,0,blend_radius_m)
  movel([0.659478, -1.258230, -2.646926, -0.807233, 1.570796, 2.230274],accel_mss,speed_ms,0,blend_radius_m)
  movel([0.659849, -1.259673, -2.646140, -0.806576, 1.570796, 2.230645],accel_mss,speed_ms,0,blend_radius_m)
  movel([0.659775, -1.263182, -2.644219, -0.804988, 1.570796, 2.230571],accel_mss,speed_ms,0,blend_radius_m)
  movel([0.659925, -1.267285, -2.641954, -0.803150, 1.570796, 2.230722],accel_mss,speed_ms,0,blend_radius_m)
  movel([0.661150, -1.272289, -2.639163, -0.800937, 1.570796, 2.231946],accel_mss,speed_ms,0,blend_radius_m)
  movel([0.662584, -1.277120, -2.636439, -0.798830, 1.570796, 2.233381],accel_mss,speed_ms,0,blend_radius_m)
  movel([0.663725, -1.282075, -2.633615, -0.796699, 1.570796, 2.234521],accel_mss,speed_ms,0,blend_radius_m)
  movel([0.664078, -1.287434, -2.630526, -0.794429, 1.570796, 2.234874],accel_mss,speed_ms,0,blend_radius_m)
  movel([0.663752, -1.290533, -2.628723, -0.793133, 1.570796, 2.234548],accel_mss,speed_ms,0,blend_radius_m)
  movel([0.663061, -1.293713, -2.626860, -0.791816, 1.570796, 2.233857],accel_mss,speed_ms,0,blend_radius_m)
  movel([0.660963, -1.300188, -2.623027, -0.789174, 1.570796, 2.231759],accel_mss,speed_ms,0,blend_radius_m)
  movel([0.658530, -1.306594, -2.619181, -0.786614, 1.570796, 2.229326],accel_mss,speed_ms,0,blend_radius_m)
  movel([0.656492, -1.312676, -2.615481, -0.784233, 1.570796, 2.227288],accel_mss,speed_ms,0,blend_radius_m)
  movel([0.654381, -1.322426, -2.609446, -0.780517, 1.570796, 2.225178],accel_mss,speed_ms,0,blend_radius_m)
  movel([0.653601, -1.326541, -2.606861, -0.778987, 1.570796, 2.224397],accel_mss,speed_ms,0,blend_radius_m)
  movel([0.652606, -1.330459, -2.604379, -0.777551, 1.570796, 2.223402],accel_mss,speed_ms,0,blend_radius_m)
  movel([0.651101, -1.334407, -2.601857, -0.776126, 1.570796, 2.221898],accel_mss,speed_ms,0,blend_radius_m)
  movel([0.648803, -1.338596, -2.599157, -0.774636, 1.570796, 2.219600],accel_mss,speed_ms,0,blend_radius_m)
  movel([0.645431, -1.343249, -2.596131, -0.773009, 1.570796, 2.216227],accel_mss,speed_ms,0,blend_radius_m)
  movel([0.640718, -1.348571, -2.592633, -0.771185, 1.570796, 2.211515],accel_mss,speed_ms,0,blend_radius_m)
  movel([0.636551, -1.352643, -2.589930, -0.769816, 1.570796, 2.207347],accel_mss,speed_ms,0,blend_radius_m)
  movel([0.632448, -1.356102, -2.587616, -0.768671, 1.570796, 2.203244],accel_mss,speed_ms,0,blend_radius_m)
  movel([0.628404, -1.358990, -2.585671, -0.767728, 1.570796, 2.199200],accel_mss,speed_ms,0,blend_radius_m)
  movel([0.624420, -1.361344, -2.584077, -0.766968, 1.570796, 2.195216],accel_mss,speed_ms,0,blend_radius_m)
  movel([0.620495, -1.363200, -2.582815, -0.766374, 1.570796, 2.191292],accel_mss,speed_ms,0,blend_radius_m)
  movel([0.616629, -1.364593, -2.581865, -0.765932, 1.570796, 2.187425],accel_mss,speed_ms,0,blend_radius_m)
  movel([0.612820, -1.365556, -2.581206, -0.765627, 1.570796, 2.183617],accel_mss,speed_ms,0,blend_radius_m)
  movel([0.609077, -1.366121, -2.580819, -0.765449, 1.570796, 2.179873],accel_mss,speed_ms,0,blend_radius_m)
  movel([0.605399, -1.366315, -2.580686, -0.765388, 1.570796, 2.176195],accel_mss,speed_ms,0,blend_radius_m)
  movel([0.601786, -1.366172, -2.580784, -0.765433, 1.570796, 2.172583],accel_mss,speed_ms,0,blend_radius_m)
  movel([0.594780, -1.364983, -2.581598, -0.765808, 1.570796, 2.165576],accel_mss,speed_ms,0,blend_radius_m)
  movel([0.588102, -1.362772, -2.583106, -0.766510, 1.570796, 2.158898],accel_mss,speed_ms,0,blend_radius_m)
  movel([0.581799, -1.359759, -2.585151, -0.767479, 1.570796, 2.152595],accel_mss,speed_ms,0,blend_radius_m)
  movel([0.576364, -1.356281, -2.587496, -0.768612, 1.570796, 2.147160],accel_mss,speed_ms,0,blend_radius_m)
  movel([0.569480, -1.351687, -2.590567, -0.770136, 1.570796, 2.140277],accel_mss,speed_ms,0,blend_radius_m)
  movel([0.561378, -1.347085, -2.593613, -0.771691, 1.570796, 2.132175],accel_mss,speed_ms,0,blend_radius_m)
  movel([0.556958, -1.345128, -2.594900, -0.772361, 1.570796, 2.127754],accel_mss,speed_ms,0,blend_radius_m)
  movel([0.552337, -1.343587, -2.595910, -0.772892, 1.570796, 2.123133],accel_mss,speed_ms,0,blend_radius_m)
  movel([0.547566, -1.342598, -2.596556, -0.773235, 1.570796, 2.118362],accel_mss,speed_ms,0,blend_radius_m)
  movel([0.542691, -1.342299, -2.596751, -0.773339, 1.570796, 2.113487],accel_mss,speed_ms,0,blend_radius_m)
  movel([0.537761, -1.342817, -2.596413, -0.773159, 1.570796, 2.108558],accel_mss,speed_ms,0,blend_radius_m)
  movel([0.532837, -1.344281, -2.595456, -0.772653, 1.570796, 2.103634],accel_mss,speed_ms,0,blend_radius_m)
  movel([0.530397, -1.345404, -2.594719, -0.772266, 1.570796, 2.101193],accel_mss,speed_ms,0,blend_radius_m)
  movel([0.527978, -1.346809, -2.593795, -0.771785, 1.570796, 2.098774],accel_mss,speed_ms,0,blend_radius_m)
  movel([0.525590, -1.348506, -2.592675, -0.771207, 1.570796, 2.096386],accel_mss,speed_ms,0,blend_radius_m)
  movel([0.523242, -1.350512, -2.591348, -0.770530, 1.570796, 2.094038],accel_mss,speed_ms,0,blend_radius_m)
  movel([0.520942, -1.352836, -2.589801, -0.769752, 1.570796, 2.091739],accel_mss,speed_ms,0,blend_radius_m)
  movel([0.518695, -1.355491, -2.588026, -0.768872, 1.570796, 2.089491],accel_mss,speed_ms,0,blend_radius_m)
  movel([0.514400, -1.361841, -2.583740, -0.766808, 1.570796, 2.085197],accel_mss,speed_ms,0,blend_radius_m)
  movel([0.513116, -1.364983, -2.581598, -0.765808, 1.570796, 2.083912],accel_mss,speed_ms,0,blend_radius_m)
  movel([0.512422, -1.368136, -2.579435, -0.764818, 1.570796, 2.083218],accel_mss,speed_ms,0,blend_radius_m)
  movel([0.512365, -1.371267, -2.577273, -0.763849, 1.570796, 2.083161],accel_mss,speed_ms,0,blend_radius_m)
  movel([0.512984, -1.374346, -2.575133, -0.762910, 1.570796, 2.083781],accel_mss,speed_ms,0,blend_radius_m)
  movel([0.516535, -1.370552, -2.577768, -0.764069, 1.570796, 2.087331],accel_mss,speed_ms,0,blend_radius_m)
  movel([0.520297, -1.367099, -2.580147, -0.765142, 1.570796, 2.091094],accel_mss,speed_ms,0,blend_radius_m)
  movel([0.524229, -1.364008, -2.582264, -0.766117, 1.570796, 2.095025],accel_mss,speed_ms,0,blend_radius_m)
  movel([0.528291, -1.361295, -2.584110, -0.766984, 1.570796, 2.099087],accel_mss,speed_ms,0,blend_radius_m)
  movel([0.532443, -1.358973, -2.585683, -0.767734, 1.570796, 2.103239],accel_mss,speed_ms,0,blend_radius_m)
  movel([0.536637, -1.357059, -2.586973, -0.768357, 1.570796, 2.107433],accel_mss,speed_ms,0,blend_radius_m)
  movel([0.540836, -1.355564, -2.587977, -0.768848, 1.570796, 2.111632],accel_mss,speed_ms,0,blend_radius_m)
  movel([0.544991, -1.354505, -2.588687, -0.769198, 1.570796, 2.115787],accel_mss,speed_ms,0,blend_radius_m)
  movel([0.549064, -1.353887, -2.589099, -0.769402, 1.570796, 2.119861],accel_mss,speed_ms,0,blend_radius_m)
  movel([0.553008, -1.353727, -2.589207, -0.769456, 1.570796, 2.123805],accel_mss,speed_ms,0,blend_radius_m)
  movel([0.556783, -1.354029, -2.589004, -0.769355, 1.570796, 2.127580],accel_mss,speed_ms,0,blend_radius_m)
  movel([0.560346, -1.354800, -2.588489, -0.769100, 1.570796, 2.131142],accel_mss,speed_ms,0,blend_radius_m)
  movel([0.563655, -1.356046, -2.587653, -0.768690, 1.570796, 2.134451],accel_mss,speed_ms,0,blend_radius_m)
  movel([0.566673, -1.357769, -2.586494, -0.768125, 1.570796, 2.137470],accel_mss,speed_ms,0,blend_radius_m)
  movel([0.569358, -1.359974, -2.585006, -0.767409, 1.570796, 2.140154],accel_mss,speed_ms,0,blend_radius_m)
  movel([0.571676, -1.362659, -2.583184, -0.766547, 1.570796, 2.142472],accel_mss,speed_ms,0,blend_radius_m)
  movel([0.573226, -1.365160, -2.581477, -0.765752, 1.570796, 2.144023],accel_mss,speed_ms,0,blend_radius_m)
  movel([0.574380, -1.367811, -2.579658, -0.764920, 1.570796, 2.145176],accel_mss,speed_ms,0,blend_radius_m)
  movel([0.575159, -1.370582, -2.577747, -0.764060, 1.570796, 2.145955],accel_mss,speed_ms,0,blend_radius_m)
  movel([0.575583, -1.373452, -2.575755, -0.763181, 1.570796, 2.146379],accel_mss,speed_ms,0,blend_radius_m)
  movel([0.575439, -1.379403, -2.571589, -0.761397, 1.570796, 2.146235],accel_mss,speed_ms,0,blend_radius_m)
  movel([0.574107, -1.385493, -2.567273, -0.759623, 1.570796, 2.144903],accel_mss,speed_ms,0,blend_radius_m)
  movel([0.571736, -1.391558, -2.562921, -0.757910, 1.570796, 2.142532],accel_mss,speed_ms,0,blend_radius_m)
  movel([0.568472, -1.397452, -2.558641, -0.756296, 1.570796, 2.139269],accel_mss,speed_ms,0,blend_radius_m)
  movel([0.564457, -1.403029, -2.554544, -0.754816, 1.570796, 2.135253],accel_mss,speed_ms,0,blend_radius_m)
  movel([0.559814, -1.408154, -2.550739, -0.753496, 1.570796, 2.130611],accel_mss,speed_ms,0,blend_radius_m)
  movel([0.554670, -1.412695, -2.547335, -0.752359, 1.570796, 2.125466],accel_mss,speed_ms,0,blend_radius_m)
  movel([0.549136, -1.416527, -2.544439, -0.751423, 1.570796, 2.119932],accel_mss,speed_ms,0,blend_radius_m)
  movel([0.543321, -1.419525, -2.542158, -0.750706, 1.570796, 2.114117],accel_mss,speed_ms,0,blend_radius_m)
  movel([0.540341, -1.420671, -2.541282, -0.750436, 1.570796, 2.111138],accel_mss,speed_ms,0,blend_radius_m)
  movel([0.537329, -1.421562, -2.540600, -0.750227, 1.570796, 2.108126],accel_mss,speed_ms,0,blend_radius_m)
  movel([0.534299, -1.422178, -2.540128, -0.750083, 1.570796, 2.105095],accel_mss,speed_ms,0,blend_radius_m)
  movel([0.531255, -1.422507, -2.539875, -0.750007, 1.570796, 2.102051],accel_mss,speed_ms,0,blend_radius_m)
  movel([0.528214, -1.422533, -2.539855, -0.750000, 1.570796, 2.099010],accel_mss,speed_ms,0,blend_radius_m)
  movel([0.525189, -1.422235, -2.540084, -0.750070, 1.570796, 2.095985],accel_mss,speed_ms,0,blend_radius_m)
  movel([0.522185, -1.421597, -2.540573, -0.750219, 1.570796, 2.092982],accel_mss,speed_ms,0,blend_radius_m)
  movel([0.519218, -1.420601, -2.541336, -0.750452, 1.570796, 2.090014],accel_mss,speed_ms,0,blend_radius_m)
  movel([0.516296, -1.419228, -2.542384, -0.750777, 1.570796, 2.087093],accel_mss,speed_ms,0,blend_radius_m)
  movel([0.513432, -1.417460, -2.543730, -0.751199, 1.570796, 2.084228],accel_mss,speed_ms,0,blend_radius_m)
  movel([0.511485, -1.415619, -2.545127, -0.751643, 1.570796, 2.082281],accel_mss,speed_ms,0,blend_radius_m)
  movel([0.506740, -1.409937, -2.549406, -0.753046, 1.570796, 2.077536],accel_mss,speed_ms,0,blend_radius_m)
  movel([0.503817, -1.405566, -2.552665, -0.754158, 1.570796, 2.074613],accel_mss,speed_ms,0,blend_radius_m)
  movel([0.500798, -1.400118, -2.556689, -0.755583, 1.570796, 2.071594],accel_mss,speed_ms,0,blend_radius_m)
  movel([0.497889, -1.393534, -2.561492, -0.757363, 1.570796, 2.068686],accel_mss,speed_ms,0,blend_radius_m)
  movel([0.495302, -1.385750, -2.567090, -0.759549, 1.570796, 2.066098],accel_mss,speed_ms,0,blend_radius_m)
  movel([0.494032, -1.379954, -2.571201, -0.761234, 1.570796, 2.064828],accel_mss,speed_ms,0,blend_radius_m)
  movel([0.493466, -1.374384, -2.575106, -0.762898, 1.570796, 2.064262],accel_mss,speed_ms,0,blend_radius_m)
  movel([0.493533, -1.369055, -2.578802, -0.764533, 1.570796, 2.064329],accel_mss,speed_ms,0,blend_radius_m)
  movel([0.494152, -1.363985, -2.582279, -0.766124, 1.570796, 2.064949],accel_mss,speed_ms,0,blend_radius_m)
  movel([0.495250, -1.359191, -2.585535, -0.767663, 1.570796, 2.066046],accel_mss,speed_ms,0,blend_radius_m)
  movel([0.496734, -1.354696, -2.588559, -0.769135, 1.570796, 2.067530],accel_mss,speed_ms,0,blend_radius_m)
  movel([0.498523, -1.350521, -2.591341, -0.770527, 1.570796, 2.069320],accel_mss,speed_ms,0,blend_radius_m)
  movel([0.500523, -1.346692, -2.593872, -0.771825, 1.570796, 2.071320],accel_mss,speed_ms,0,blend_radius_m)
  movel([0.504798, -1.340159, -2.598144, -0.774086, 1.570796, 2.075595],accel_mss,speed_ms,0,blend_radius_m)
  movel([0.508802, -1.335286, -2.601292, -0.775811, 1.570796, 2.079599],accel_mss,speed_ms,0,blend_radius_m)
  movel([0.511766, -1.332247, -2.603239, -0.776903, 1.570796, 2.082563],accel_mss,speed_ms,0,blend_radius_m)
  movel([0.512921, -1.331202, -2.603906, -0.777281, 1.570796, 2.083717],accel_mss,speed_ms,0,blend_radius_m)
  movel([0.518608, -1.326597, -2.606826, -0.778966, 1.570796, 2.089405],accel_mss,speed_ms,0,blend_radius_m)
  movel([0.524249, -1.322741, -2.609249, -0.780399, 1.570796, 2.095046],accel_mss,speed_ms,0,blend_radius_m)
  movel([0.529796, -1.319587, -2.611216, -0.781586, 1.570796, 2.100593],accel_mss,speed_ms,0,blend_radius_m)
  movel([0.535212, -1.317091, -2.612764, -0.782535, 1.570796, 2.106008],accel_mss,speed_ms,0,blend_radius_m)
  movel([0.540452, -1.315195, -2.613933, -0.783260, 1.570796, 2.111249],accel_mss,speed_ms,0,blend_radius_m)
  movel([0.545478, -1.313849, -2.614761, -0.783779, 1.570796, 2.116274],accel_mss,speed_ms,0,blend_radius_m)
  movel([0.550257, -1.312989, -2.615288, -0.784111, 1.570796, 2.121054],accel_mss,speed_ms,0,blend_radius_m)
  movel([0.554752, -1.312557, -2.615554, -0.784279, 1.570796, 2.125548],accel_mss,speed_ms,0,blend_radius_m)
  movel([0.562766, -1.312710, -2.615459, -0.784219, 1.570796, 2.133562],accel_mss,speed_ms,0,blend_radius_m)
  movel([0.569299, -1.313774, -2.614807, -0.783808, 1.570796, 2.140095],accel_mss,speed_ms,0,blend_radius_m)
  movel([0.574149, -1.315209, -2.613925, -0.783255, 1.570796, 2.144945],accel_mss,speed_ms,0,blend_radius_m)
  movel([0.577138, -1.316464, -2.613151, -0.782774, 1.570796, 2.147934],accel_mss,speed_ms,0,blend_radius_m)
  movel([0.584260, -1.319385, -2.611341, -0.781662, 1.570796, 2.155057],accel_mss,speed_ms,0,blend_radius_m)
  movel([0.591498, -1.323204, -2.608959, -0.780226, 1.570796, 2.162294],accel_mss,speed_ms,0,blend_radius_m)
  movel([0.598673, -1.327314, -2.606373, -0.778702, 1.570796, 2.169469],accel_mss,speed_ms,0,blend_radius_m)
  movel([0.605633, -1.331116, -2.603960, -0.777312, 1.570796, 2.176429],accel_mss,speed_ms,0,blend_radius_m)
  movel([0.612253, -1.334006, -2.602114, -0.776269, 1.570796, 2.183050],accel_mss,speed_ms,0,blend_radius_m)
  movel([0.615400, -1.334920, -2.601527, -0.775942, 1.570796, 2.186196],accel_mss,speed_ms,0,blend_radius_m)
  movel([0.618423, -1.335377, -2.601234, -0.775778, 1.570796, 2.189219],accel_mss,speed_ms,0,blend_radius_m)
  movel([0.621310, -1.335301, -2.601283, -0.775806, 1.570796, 2.192106],accel_mss,speed_ms,0,blend_radius_m)
  movel([0.624052, -1.334610, -2.601726, -0.776053, 1.570796, 2.194848],accel_mss,speed_ms,0,blend_radius_m)
  movel([0.626639, -1.333228, -2.602612, -0.776549, 1.570796, 2.197436],accel_mss,speed_ms,0,blend_radius_m)
  movel([0.629060, -1.331068, -2.603991, -0.777330, 1.570796, 2.199856],accel_mss,speed_ms,0,blend_radius_m)
  movel([0.630565, -1.329194, -2.605183, -0.778013, 1.570796, 2.201361],accel_mss,speed_ms,0,blend_radius_m)
  movel([0.631712, -1.327310, -2.606375, -0.778703, 1.570796, 2.202508],accel_mss,speed_ms,0,blend_radius_m)
  movel([0.633073, -1.323534, -2.608752, -0.780103, 1.570796, 2.203870],accel_mss,speed_ms,0,blend_radius_m)
  movel([0.633420, -1.319757, -2.611111, -0.781522, 1.570796, 2.204216],accel_mss,speed_ms,0,blend_radius_m)
  movel([0.633018, -1.316013, -2.613429, -0.782947, 1.570796, 2.203815],accel_mss,speed_ms,0,blend_radius_m)
  movel([0.631109, -1.308726, -2.617889, -0.785773, 1.570796, 2.201905],accel_mss,speed_ms,0,blend_radius_m)
  movel([0.630172, -1.305236, -2.620001, -0.787152, 1.570796, 2.200968],accel_mss,speed_ms,0,blend_radius_m)
  movel([0.629643, -1.301878, -2.622018, -0.788494, 1.570796, 2.200439],accel_mss,speed_ms,0,blend_radius_m)
  movel([0.629911, -1.296386, -2.625284, -0.790719, 1.570796, 2.200707],accel_mss,speed_ms,0,blend_radius_m)
  movel([0.631145, -1.289408, -2.629379, -0.793602, 1.570796, 2.201942],accel_mss,speed_ms,0,blend_radius_m)
  movel([0.633069, -1.282195, -2.633546, -0.796648, 1.570796, 2.203865],accel_mss,speed_ms,0,blend_radius_m)
  movel([0.635383, -1.276056, -2.637041, -0.799291, 1.570796, 2.206179],accel_mss,speed_ms,0,blend_radius_m)
  movel([0.637598, -1.272263, -2.639177, -0.800948, 1.570796, 2.208394],accel_mss,speed_ms,0,blend_radius_m)
  movel([0.640692, -1.267665, -2.641743, -0.802981, 1.570796, 2.211489],accel_mss,speed_ms,0,blend_radius_m)
  movel([0.643604, -1.263273, -2.644169, -0.804947, 1.570796, 2.214400],accel_mss,speed_ms,0,blend_radius_m)
  movel([0.645246, -1.260124, -2.645894, -0.806371, 1.570796, 2.216042],accel_mss,speed_ms,0,blend_radius_m)
  movel([0.645630, -1.256942, -2.647625, -0.807822, 1.570796, 2.216427],accel_mss,speed_ms,0,blend_radius_m)
  movel([0.645451, -1.253334, -2.649573, -0.809482, 1.570796, 2.216247],accel_mss,speed_ms,0,blend_radius_m)
  movel([0.645306, -1.249287, -2.651739, -0.811363, 1.570796, 2.216102],accel_mss,speed_ms,0,blend_radius_m)
  movel([0.645820, -1.244779, -2.654129, -0.813482, 1.570796, 2.216616],accel_mss,speed_ms,0,blend_radius_m)
  movel([0.646760, -1.241987, -2.655596, -0.814805, 1.570796, 2.217556],accel_mss,speed_ms,0,blend_radius_m)
  speed_ms = 0.003
  movel([0.646760, -1.234835, -2.652122, -0.825432, 1.570796, 2.217556],accel_mss,speed_ms,0,blend_radius_m)
  speed_ms = 0.03
  movel([0.646760, -1.207578, -2.637954, -0.866856, 1.570796, 2.217556],accel_mss,speed_ms,0,blend_radius_m)
  #M_RunCode9
  movel([0.495863, -1.322864, -2.572500, -0.817025, 1.570796, 2.066659],accel_mss,speed_ms,0,blend_radius_m)
  #M_RunCode3
  movel([0.495863, -1.348500, -2.585150, -0.778739, 1.570796, 2.066659],accel_mss,speed_ms,0,blend_radius_m)
  speed_ms = 0.003
  movel([0.495863, -1.355171, -2.588241, -0.768978, 1.570796, 2.066659],accel_mss,speed_ms,0,blend_radius_m)
  speed_ms = 0.007
  movel([0.488256, -1.353194, -2.589562, -0.769633, 1.570796, 2.059052],accel_mss,speed_ms,0,blend_radius_m)
  movel([0.480522, -1.352226, -2.590208, -0.769955, 1.570796, 2.051318],accel_mss,speed_ms,0,blend_radius_m)
  movel([0.472764, -1.352148, -2.590260, -0.769981, 1.570796, 2.043561],accel_mss,speed_ms,0,blend_radius_m)
  movel([0.465081, -1.352836, -2.589801, -0.769752, 1.570796, 2.035877],accel_mss,speed_ms,0,blend_radius_m)
  movel([0.457570, -1.354169, -2.588911, -0.769309, 1.570796, 2.028366],accel_mss,speed_ms,0,blend_radius_m)
  movel([0.450325, -1.356016, -2.587674, -0.768699, 1.570796, 2.021121],accel_mss,speed_ms,0,blend_radius_m)
  movel([0.443427, -1.358256, -2.586167, -0.767967, 1.570796, 2.014223],accel_mss,speed_ms,0,blend_radius_m)
  movel([0.436964, -1.360758, -2.584475, -0.767156, 1.570796, 2.007760],accel_mss,speed_ms,0,blend_radius_m)
  movel([0.431009, -1.363400, -2.582678, -0.766310, 1.570796, 2.001805],accel_mss,speed_ms,0,blend_radius_m)
  movel([0.425637, -1.366063, -2.580859, -0.765467, 1.570796, 1.996433],accel_mss,speed_ms,0,blend_radius_m)
  movel([0.416915, -1.370970, -2.577478, -0.763941, 1.570796, 1.987711],accel_mss,speed_ms,0,blend_radius_m)
  movel([0.411311, -1.374565, -2.574980, -0.762844, 1.570796, 1.982108],accel_mss,speed_ms,0,blend_radius_m)
  movel([0.409332, -1.375956, -2.574008, -0.762424, 1.570796, 1.980128],accel_mss,speed_ms,0,blend_radius_m)
  movel([0.406132, -1.378070, -2.572527, -0.761792, 1.570796, 1.976928],accel_mss,speed_ms,0,blend_radius_m)
  movel([0.398032, -1.384142, -2.568235, -0.760012, 1.570796, 1.968828],accel_mss,speed_ms,0,blend_radius_m)
  movel([0.392858, -1.388526, -2.565103, -0.758760, 1.570796, 1.963654],accel_mss,speed_ms,0,blend_radius_m)
  movel([0.387316, -1.393722, -2.561355, -0.757311, 1.570796, 1.958112],accel_mss,speed_ms,0,blend_radius_m)
  movel([0.381690, -1.399664, -2.557022, -0.755704, 1.570796, 1.952486],accel_mss,speed_ms,0,blend_radius_m)
  movel([0.376259, -1.406282, -2.552133, -0.753974, 1.570796, 1.947055],accel_mss,speed_ms,0,blend_radius_m)
  movel([0.371293, -1.413499, -2.546729, -0.752161, 1.570796, 1.942089],accel_mss,speed_ms,0,blend_radius_m)
  movel([0.367051, -1.421246, -2.540842, -0.750301, 1.570796, 1.937847],accel_mss,speed_ms,0,blend_radius_m)
  movel([0.365277, -1.425297, -2.537728, -0.749364, 1.570796, 1.936074],accel_mss,speed_ms,0,blend_radius_m)
  movel([0.363779, -1.429454, -2.534507, -0.748428, 1.570796, 1.934575],accel_mss,speed_ms,0,blend_radius_m)
  movel([0.362580, -1.433709, -2.531182, -0.747497, 1.570796, 1.933376],accel_mss,speed_ms,0,blend_radius_m)
  movel([0.361710, -1.438058, -2.527757, -0.746575, 1.570796, 1.932506],accel_mss,speed_ms,0,blend_radius_m)
  movel([0.361197, -1.442491, -2.524235, -0.745663, 1.570796, 1.931993],accel_mss,speed_ms,0,blend_radius_m)
  movel([0.361065, -1.447004, -2.520619, -0.744766, 1.570796, 1.931862],accel_mss,speed_ms,0,blend_radius_m)
  movel([0.361342, -1.451590, -2.516912, -0.743886, 1.570796, 1.932138],accel_mss,speed_ms,0,blend_radius_m)
  movel([0.362047, -1.456247, -2.513116, -0.743026, 1.570796, 1.932843],accel_mss,speed_ms,0,blend_radius_m)
  movel([0.363206, -1.460972, -2.509229, -0.742187, 1.570796, 1.934003],accel_mss,speed_ms,0,blend_radius_m)
  movel([0.364840, -1.465760, -2.505257, -0.741372, 1.570796, 1.935636],accel_mss,speed_ms,0,blend_radius_m)
  movel([0.366967, -1.470612, -2.501194, -0.740583, 1.570796, 1.937763],accel_mss,speed_ms,0,blend_radius_m)
  movel([0.369612, -1.475526, -2.497042, -0.739821, 1.570796, 1.940409],accel_mss,speed_ms,0,blend_radius_m)
  movel([0.369849, -1.475889, -2.496734, -0.739766, 1.570796, 1.940645],accel_mss,speed_ms,0,blend_radius_m)
  movel([0.373245, -1.480255, -2.493011, -0.739123, 1.570796, 1.944041],accel_mss,speed_ms,0,blend_radius_m)
  movel([0.376738, -1.484085, -2.489721, -0.738583, 1.570796, 1.947534],accel_mss,speed_ms,0,blend_radius_m)
  movel([0.380316, -1.487407, -2.486848, -0.738133, 1.570796, 1.951113],accel_mss,speed_ms,0,blend_radius_m)
  movel([0.383970, -1.490259, -2.484369, -0.737761, 1.570796, 1.954766],accel_mss,speed_ms,0,blend_radius_m)
  movel([0.387689, -1.492665, -2.482266, -0.737457, 1.570796, 1.958485],accel_mss,speed_ms,0,blend_radius_m)
  movel([0.391463, -1.494657, -2.480519, -0.737212, 1.570796, 1.962259],accel_mss,speed_ms,0,blend_radius_m)
  movel([0.395275, -1.496263, -2.479106, -0.737020, 1.570796, 1.966071],accel_mss,speed_ms,0,blend_radius_m)
  movel([0.399119, -1.497509, -2.478007, -0.736873, 1.570796, 1.969916],accel_mss,speed_ms,0,blend_radius_m)
  movel([0.402982, -1.498422, -2.477200, -0.736767, 1.570796, 1.973779],accel_mss,speed_ms,0,blend_radius_m)
  movel([0.406855, -1.499024, -2.476667, -0.736698, 1.570796, 1.977651],accel_mss,speed_ms,0,blend_radius_m)
  movel([0.410720, -1.499343, -2.476385, -0.736661, 1.570796, 1.981517],accel_mss,speed_ms,0,blend_radius_m)
  movel([0.414570, -1.499401, -2.476333, -0.736655, 1.570796, 1.985366],accel_mss,speed_ms,0,blend_radius_m)
  movel([0.422160, -1.498835, -2.476834, -0.736719, 1.570796, 1.992957],accel_mss,speed_ms,0,blend_radius_m)
  movel([0.429524, -1.497515, -2.478002, -0.736872, 1.570796, 2.000320],accel_mss,speed_ms,0,blend_radius_m)
  movel([0.436538, -1.495628, -2.479665, -0.737095, 1.570796, 2.007334],accel_mss,speed_ms,0,blend_radius_m)
  movel([0.443082, -1.493362, -2.481656, -0.737371, 1.570796, 2.013879],accel_mss,speed_ms,0,blend_radius_m)
  movel([0.449022, -1.490905, -2.483805, -0.737679, 1.570796, 2.019818],accel_mss,speed_ms,0,blend_radius_m)
  movel([0.454218, -1.488450, -2.485944, -0.737996, 1.570796, 2.025014],accel_mss,speed_ms,0,blend_radius_m)
  movel([0.461790, -1.484327, -2.489512, -0.738550, 1.570796, 2.032587],accel_mss,speed_ms,0,blend_radius_m)
  movel([0.464584, -1.482592, -2.491006, -0.738791, 1.570796, 2.035380],accel_mss,speed_ms,0,blend_radius_m)
  movel([0.466299, -1.481588, -2.491869, -0.738932, 1.570796, 2.037095],accel_mss,speed_ms,0,blend_radius_m)
  movel([0.470942, -1.478624, -2.494405, -0.739359, 1.570796, 2.041738],accel_mss,speed_ms,0,blend_radius_m)
  movel([0.477785, -1.473756, -2.498542, -0.740091, 1.570796, 2.048581],accel_mss,speed_ms,0,blend_radius_m)
  movel([0.486114, -1.467025, -2.504201, -0.741163, 1.570796, 2.056910],accel_mss,speed_ms,0,blend_radius_m)
  movel([0.490613, -1.462965, -2.507580, -0.741844, 1.570796, 2.061409],accel_mss,speed_ms,0,blend_radius_m)
  movel([0.495218, -1.458441, -2.511316, -0.742632, 1.570796, 2.066015],accel_mss,speed_ms,0,blend_radius_m)
  movel([0.499837, -1.453451, -2.515400, -0.743539, 1.570796, 2.070633],accel_mss,speed_ms,0,blend_radius_m)
  movel([0.504380, -1.447988, -2.519827, -0.744575, 1.570796, 2.075176],accel_mss,speed_ms,0,blend_radius_m)
  movel([0.508749, -1.442046, -2.524590, -0.745753, 1.570796, 2.079546],accel_mss,speed_ms,0,blend_radius_m)
  movel([0.512852, -1.435616, -2.529684, -0.747089, 1.570796, 2.083648],accel_mss,speed_ms,0,blend_radius_m)
  movel([0.516586, -1.428690, -2.535100, -0.748598, 1.570796, 2.087382],accel_mss,speed_ms,0,blend_radius_m)
  movel([0.519848, -1.421256, -2.540835, -0.750299, 1.570796, 2.090644],accel_mss,speed_ms,0,blend_radius_m)
  speed_ms = 0.003
  movel([0.519848, -1.414938, -2.537960, -0.759491, 1.570796, 2.090644],accel_mss,speed_ms,0,blend_radius_m)
  speed_ms = 0.03
  movel([0.519848, -1.390554, -2.526171, -0.795665, 1.570796, 2.090644],accel_mss,speed_ms,0,blend_radius_m)
  #M_RunCode9
  movel([0.488485, -1.382321, -2.532140, -0.797927, 1.570796, 2.059282],accel_mss,speed_ms,0,blend_radius_m)
  #M_RunCode3
